REGION Network 5: 外呼下面有目标
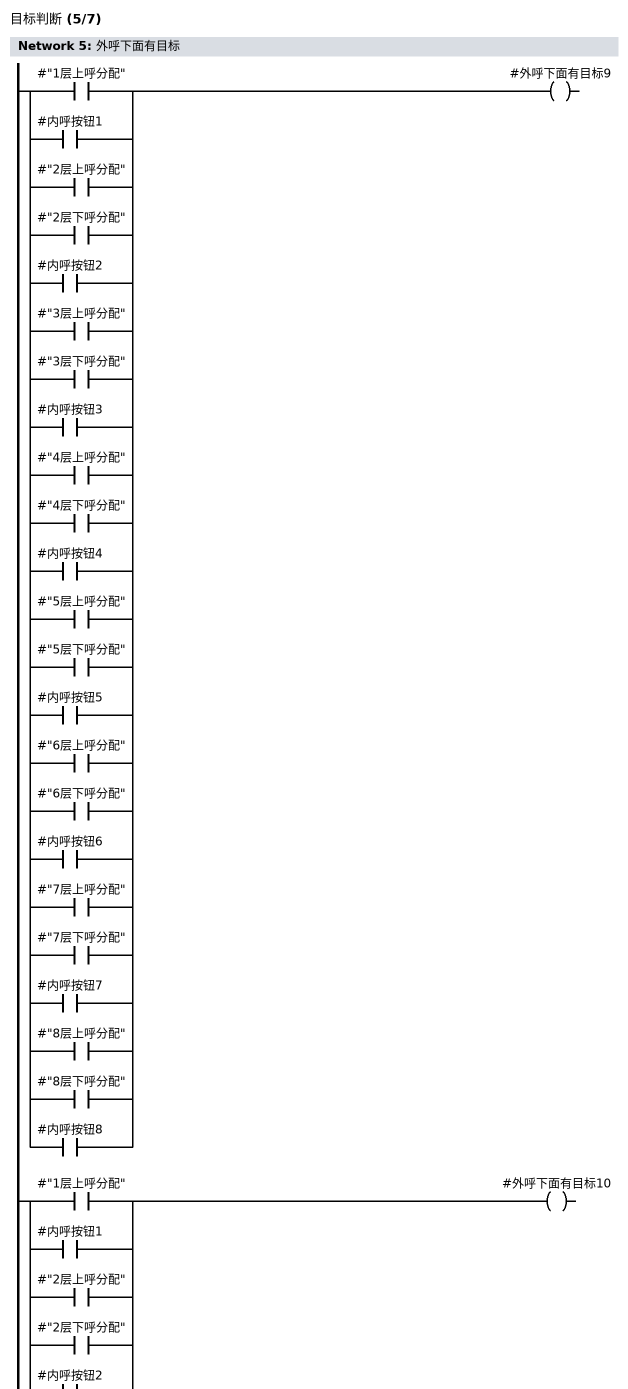
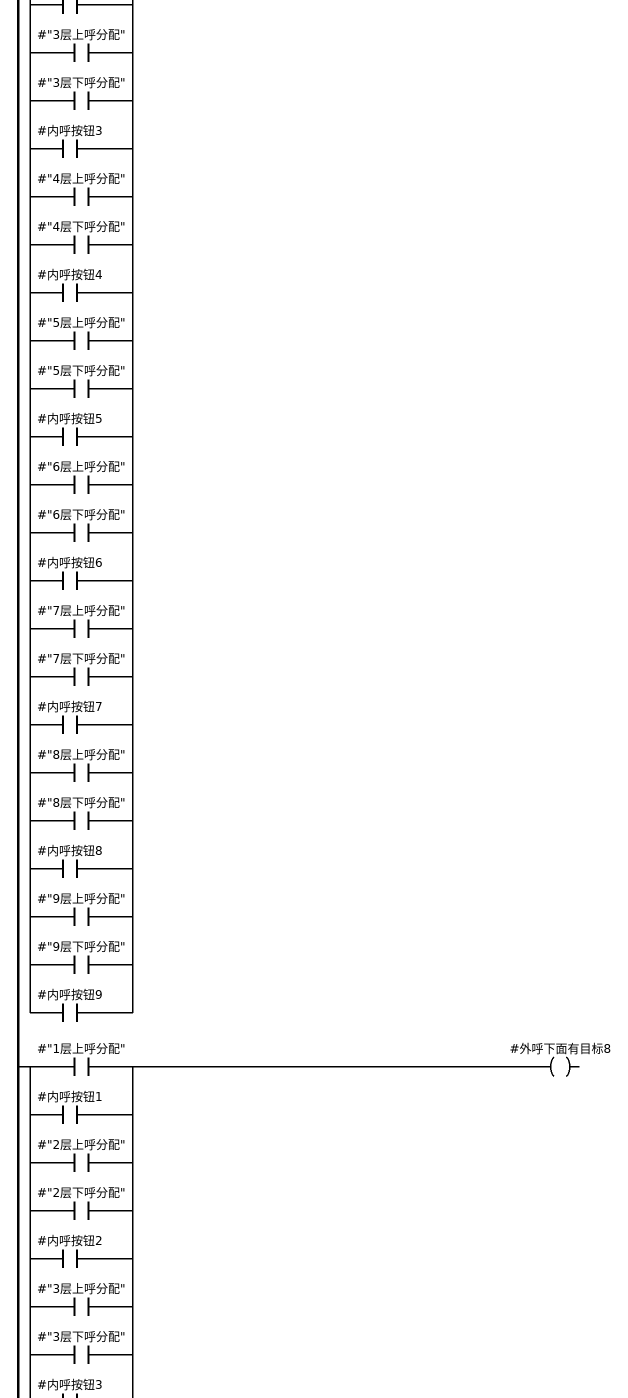
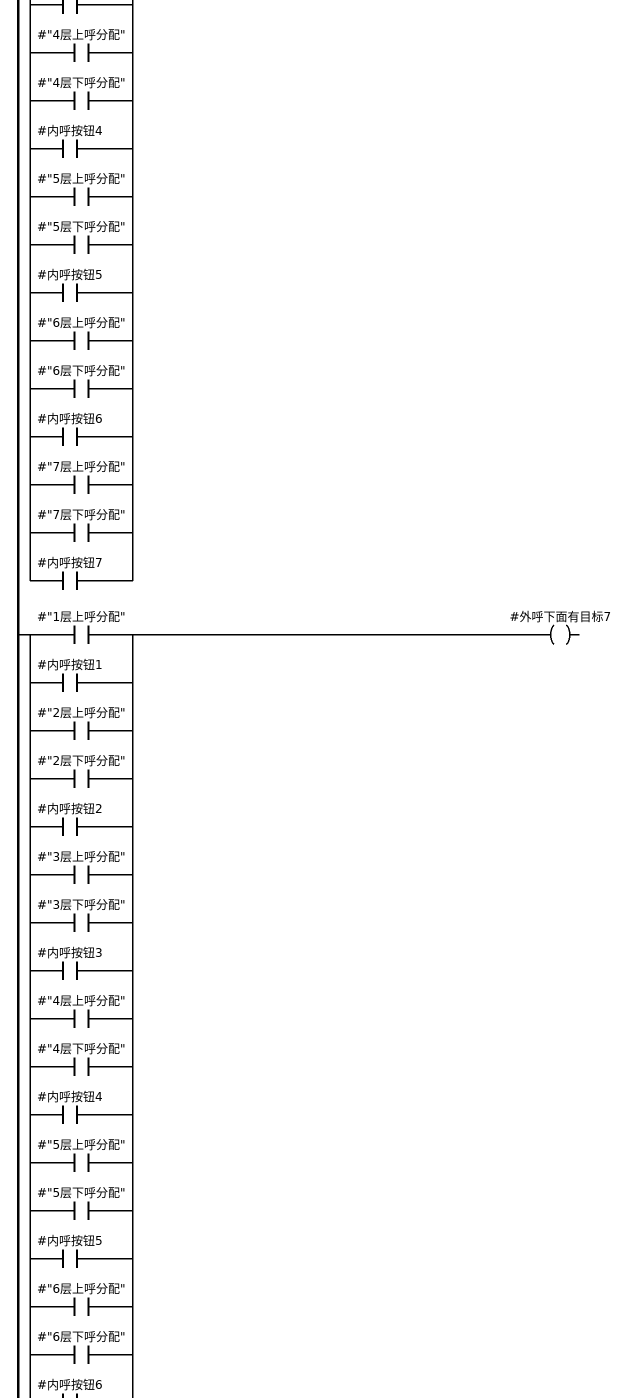
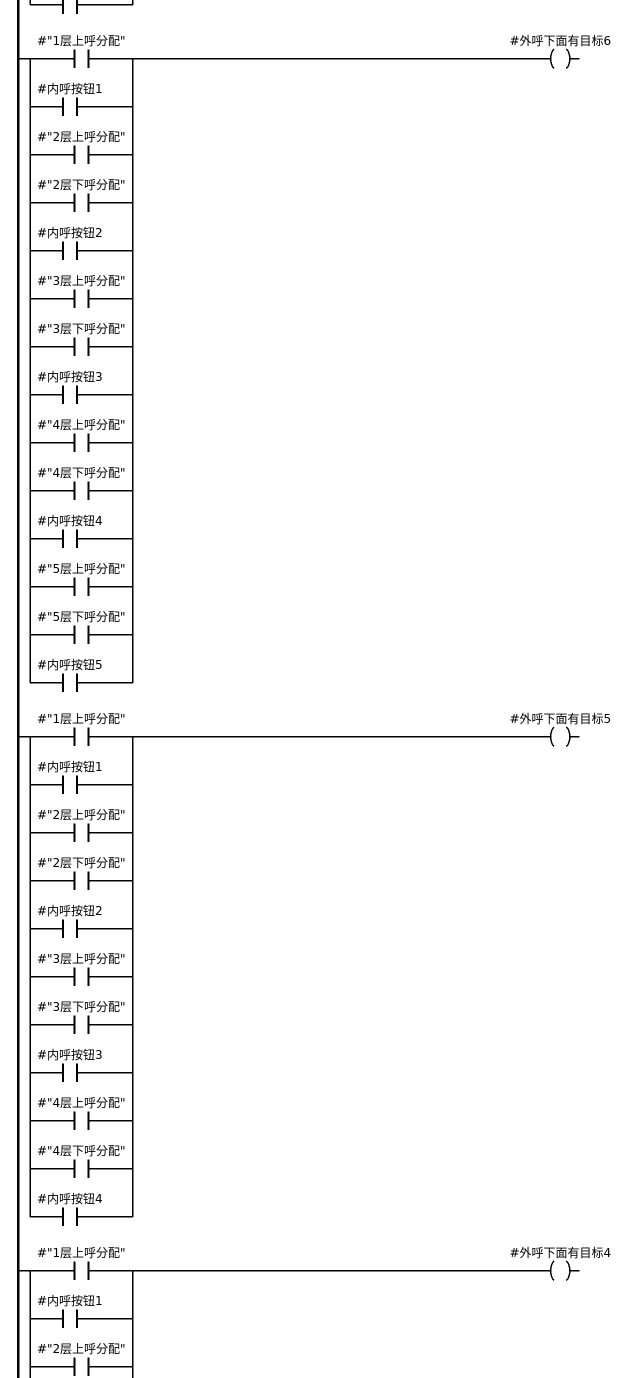
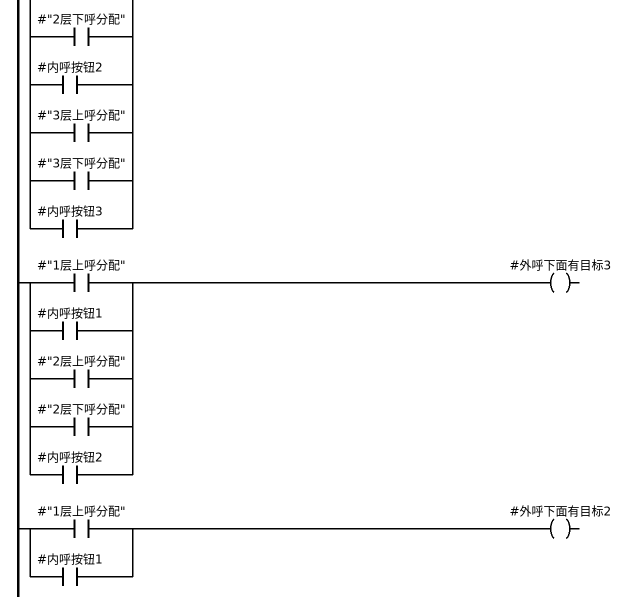
   RUNG wire#powerrail
      Contact( #"1层上呼分配" )
      wire#w1
      Coil( #外呼下面有目标9 )
   END_RUNG
   RUNG wire#powerrail
      Contact( #内呼按钮1 )
   END_RUNG wire#w1
   RUNG wire#powerrail
      Contact( #"2层上呼分配" )
   END_RUNG wire#w1
   RUNG wire#powerrail
      Contact( #"2层下呼分配" )
   END_RUNG wire#w1
   RUNG wire#powerrail
      Contact( #内呼按钮2 )
   END_RUNG wire#w1
   RUNG wire#powerrail
      Contact( #"3层上呼分配" )
   END_RUNG wire#w1
   RUNG wire#powerrail
      Contact( #"3层下呼分配" )
   END_RUNG wire#w1
   RUNG wire#powerrail
      Contact( #内呼按钮3 )
   END_RUNG wire#w1
   RUNG wire#powerrail
      Contact( #"4层上呼分配" )
   END_RUNG wire#w1
   RUNG wire#powerrail
      Contact( #"4层下呼分配" )
   END_RUNG wire#w1
   RUNG wire#powerrail
      Contact( #内呼按钮4 )
   END_RUNG wire#w1
   RUNG wire#powerrail
      Contact( #"5层上呼分配" )
   END_RUNG wire#w1
   RUNG wire#powerrail
      Contact( #"5层下呼分配" )
   END_RUNG wire#w1
   RUNG wire#powerrail
      Contact( #内呼按钮5 )
   END_RUNG wire#w1
   RUNG wire#powerrail
      Contact( #"6层上呼分配" )
   END_RUNG wire#w1
   RUNG wire#powerrail
      Contact( #"6层下呼分配" )
   END_RUNG wire#w1
   RUNG wire#powerrail
      Contact( #内呼按钮6 )
   END_RUNG wire#w1
   RUNG wire#powerrail
      Contact( #"7层上呼分配" )
   END_RUNG wire#w1
   RUNG wire#powerrail
      Contact( #"7层下呼分配" )
   END_RUNG wire#w1
   RUNG wire#powerrail
      Contact( #内呼按钮7 )
   END_RUNG wire#w1
   RUNG wire#powerrail
      Contact( #"8层上呼分配" )
   END_RUNG wire#w1
   RUNG wire#powerrail
      Contact( #"8层下呼分配" )
   END_RUNG wire#w1
   RUNG wire#powerrail
      Contact( #内呼按钮8 )
   END_RUNG wire#w1
   RUNG wire#powerrail
      Contact( #"1层上呼分配" )
      wire#w2
      Coil( #外呼下面有目标10 )
   END_RUNG
   RUNG wire#powerrail
      Contact( #内呼按钮1 )
   END_RUNG wire#w2
   RUNG wire#powerrail
      Contact( #"2层上呼分配" )
   END_RUNG wire#w2
   RUNG wire#powerrail
      Contact( #"2层下呼分配" )
   END_RUNG wire#w2
   RUNG wire#powerrail
      Contact( #内呼按钮2 )
   END_RUNG wire#w2
   RUNG wire#powerrail
      Contact( #"3层上呼分配" )
   END_RUNG wire#w2
   RUNG wire#powerrail
      Contact( #"3层下呼分配" )
   END_RUNG wire#w2
   RUNG wire#powerrail
      Contact( #内呼按钮3 )
   END_RUNG wire#w2
   RUNG wire#powerrail
      Contact( #"4层上呼分配" )
   END_RUNG wire#w2
   RUNG wire#powerrail
      Contact( #"4层下呼分配" )
   END_RUNG wire#w2
   RUNG wire#powerrail
      Contact( #内呼按钮4 )
   END_RUNG wire#w2
   RUNG wire#powerrail
      Contact( #"5层上呼分配" )
   END_RUNG wire#w2
   RUNG wire#powerrail
      Contact( #"5层下呼分配" )
   END_RUNG wire#w2
   RUNG wire#powerrail
      Contact( #内呼按钮5 )
   END_RUNG wire#w2
   RUNG wire#powerrail
      Contact( #"6层上呼分配" )
   END_RUNG wire#w2
   RUNG wire#powerrail
      Contact( #"6层下呼分配" )
   END_RUNG wire#w2
   RUNG wire#powerrail
      Contact( #内呼按钮6 )
   END_RUNG wire#w2
   RUNG wire#powerrail
      Contact( #"7层上呼分配" )
   END_RUNG wire#w2
   RUNG wire#powerrail
      Contact( #"7层下呼分配" )
   END_RUNG wire#w2
   RUNG wire#powerrail
      Contact( #内呼按钮7 )
   END_RUNG wire#w2
   RUNG wire#powerrail
      Contact( #"8层上呼分配" )
   END_RUNG wire#w2
   RUNG wire#powerrail
      Contact( #"8层下呼分配" )
   END_RUNG wire#w2
   RUNG wire#powerrail
      Contact( #内呼按钮8 )
   END_RUNG wire#w2
   RUNG wire#powerrail
      Contact( #"9层上呼分配" )
   END_RUNG wire#w2
   RUNG wire#powerrail
      Contact( #"9层下呼分配" )
   END_RUNG wire#w2
   RUNG wire#powerrail
      Contact( #内呼按钮9 )
   END_RUNG wire#w2
   RUNG wire#powerrail
      Contact( #"1层上呼分配" )
      wire#w3
      Coil( #外呼下面有目标8 )
   END_RUNG
   RUNG wire#powerrail
      Contact( #内呼按钮1 )
   END_RUNG wire#w3
   RUNG wire#powerrail
      Contact( #"2层上呼分配" )
   END_RUNG wire#w3
   RUNG wire#powerrail
      Contact( #"2层下呼分配" )
   END_RUNG wire#w3
   RUNG wire#powerrail
      Contact( #内呼按钮2 )
   END_RUNG wire#w3
   RUNG wire#powerrail
      Contact( #"3层上呼分配" )
   END_RUNG wire#w3
   RUNG wire#powerrail
      Contact( #"3层下呼分配" )
   END_RUNG wire#w3
   RUNG wire#powerrail
      Contact( #内呼按钮3 )
   END_RUNG wire#w3
   RUNG wire#powerrail
      Contact( #"4层上呼分配" )
   END_RUNG wire#w3
   RUNG wire#powerrail
      Contact( #"4层下呼分配" )
   END_RUNG wire#w3
   RUNG wire#powerrail
      Contact( #内呼按钮4 )
   END_RUNG wire#w3
   RUNG wire#powerrail
      Contact( #"5层上呼分配" )
   END_RUNG wire#w3
   RUNG wire#powerrail
      Contact( #"5层下呼分配" )
   END_RUNG wire#w3
   RUNG wire#powerrail
      Contact( #内呼按钮5 )
   END_RUNG wire#w3
   RUNG wire#powerrail
      Contact( #"6层上呼分配" )
   END_RUNG wire#w3
   RUNG wire#powerrail
      Contact( #"6层下呼分配" )
   END_RUNG wire#w3
   RUNG wire#powerrail
      Contact( #内呼按钮6 )
   END_RUNG wire#w3
   RUNG wire#powerrail
      Contact( #"7层上呼分配" )
   END_RUNG wire#w3
   RUNG wire#powerrail
      Contact( #"7层下呼分配" )
   END_RUNG wire#w3
   RUNG wire#powerrail
      Contact( #内呼按钮7 )
   END_RUNG wire#w3
   RUNG wire#powerrail
      Contact( #"1层上呼分配" )
      wire#w4
      Coil( #外呼下面有目标7 )
   END_RUNG
   RUNG wire#powerrail
      Contact( #内呼按钮1 )
   END_RUNG wire#w4
   RUNG wire#powerrail
      Contact( #"2层上呼分配" )
   END_RUNG wire#w4
   RUNG wire#powerrail
      Contact( #"2层下呼分配" )
   END_RUNG wire#w4
   RUNG wire#powerrail
      Contact( #内呼按钮2 )
   END_RUNG wire#w4
   RUNG wire#powerrail
      Contact( #"3层上呼分配" )
   END_RUNG wire#w4
   RUNG wire#powerrail
      Contact( #"3层下呼分配" )
   END_RUNG wire#w4
   RUNG wire#powerrail
      Contact( #内呼按钮3 )
   END_RUNG wire#w4
   RUNG wire#powerrail
      Contact( #"4层上呼分配" )
   END_RUNG wire#w4
   RUNG wire#powerrail
      Contact( #"4层下呼分配" )
   END_RUNG wire#w4
   RUNG wire#powerrail
      Contact( #内呼按钮4 )
   END_RUNG wire#w4
   RUNG wire#powerrail
      Contact( #"5层上呼分配" )
   END_RUNG wire#w4
   RUNG wire#powerrail
      Contact( #"5层下呼分配" )
   END_RUNG wire#w4
   RUNG wire#powerrail
      Contact( #内呼按钮5 )
   END_RUNG wire#w4
   RUNG wire#powerrail
      Contact( #"6层上呼分配" )
   END_RUNG wire#w4
   RUNG wire#powerrail
      Contact( #"6层下呼分配" )
   END_RUNG wire#w4
   RUNG wire#powerrail
      Contact( #内呼按钮6 )
   END_RUNG wire#w4
   RUNG wire#powerrail
      Contact( #"1层上呼分配" )
      wire#w5
      Coil( #外呼下面有目标6 )
   END_RUNG
   RUNG wire#powerrail
      Contact( #内呼按钮1 )
   END_RUNG wire#w5
   RUNG wire#powerrail
      Contact( #"2层上呼分配" )
   END_RUNG wire#w5
   RUNG wire#powerrail
      Contact( #"2层下呼分配" )
   END_RUNG wire#w5
   RUNG wire#powerrail
      Contact( #内呼按钮2 )
   END_RUNG wire#w5
   RUNG wire#powerrail
      Contact( #"3层上呼分配" )
   END_RUNG wire#w5
   RUNG wire#powerrail
      Contact( #"3层下呼分配" )
   END_RUNG wire#w5
   RUNG wire#powerrail
      Contact( #内呼按钮3 )
   END_RUNG wire#w5
   RUNG wire#powerrail
      Contact( #"4层上呼分配" )
   END_RUNG wire#w5
   RUNG wire#powerrail
      Contact( #"4层下呼分配" )
   END_RUNG wire#w5
   RUNG wire#powerrail
      Contact( #内呼按钮4 )
   END_RUNG wire#w5
   RUNG wire#powerrail
      Contact( #"5层上呼分配" )
   END_RUNG wire#w5
   RUNG wire#powerrail
      Contact( #"5层下呼分配" )
   END_RUNG wire#w5
   RUNG wire#powerrail
      Contact( #内呼按钮5 )
   END_RUNG wire#w5
   RUNG wire#powerrail
      Contact( #"1层上呼分配" )
      wire#w6
      Coil( #外呼下面有目标5 )
   END_RUNG
   RUNG wire#powerrail
      Contact( #内呼按钮1 )
   END_RUNG wire#w6
   RUNG wire#powerrail
      Contact( #"2层上呼分配" )
   END_RUNG wire#w6
   RUNG wire#powerrail
      Contact( #"2层下呼分配" )
   END_RUNG wire#w6
   RUNG wire#powerrail
      Contact( #内呼按钮2 )
   END_RUNG wire#w6
   RUNG wire#powerrail
      Contact( #"3层上呼分配" )
   END_RUNG wire#w6
   RUNG wire#powerrail
      Contact( #"3层下呼分配" )
   END_RUNG wire#w6
   RUNG wire#powerrail
      Contact( #内呼按钮3 )
   END_RUNG wire#w6
   RUNG wire#powerrail
      Contact( #"4层上呼分配" )
   END_RUNG wire#w6
   RUNG wire#powerrail
      Contact( #"4层下呼分配" )
   END_RUNG wire#w6
   RUNG wire#powerrail
      Contact( #内呼按钮4 )
   END_RUNG wire#w6
   RUNG wire#powerrail
      Contact( #"1层上呼分配" )
      wire#w7
      Coil( #外呼下面有目标4 )
   END_RUNG
   RUNG wire#powerrail
      Contact( #内呼按钮1 )
   END_RUNG wire#w7
   RUNG wire#powerrail
      Contact( #"2层上呼分配" )
   END_RUNG wire#w7
   RUNG wire#powerrail
      Contact( #"2层下呼分配" )
   END_RUNG wire#w7
   RUNG wire#powerrail
      Contact( #内呼按钮2 )
   END_RUNG wire#w7
   RUNG wire#powerrail
      Contact( #"3层上呼分配" )
   END_RUNG wire#w7
   RUNG wire#powerrail
      Contact( #"3层下呼分配" )
   END_RUNG wire#w7
   RUNG wire#powerrail
      Contact( #内呼按钮3 )
   END_RUNG wire#w7
   RUNG wire#powerrail
      Contact( #"1层上呼分配" )
      wire#w8
      Coil( #外呼下面有目标3 )
   END_RUNG
   RUNG wire#powerrail
      Contact( #内呼按钮1 )
   END_RUNG wire#w8
   RUNG wire#powerrail
      Contact( #"2层上呼分配" )
   END_RUNG wire#w8
   RUNG wire#powerrail
      Contact( #"2层下呼分配" )
   END_RUNG wire#w8
   RUNG wire#powerrail
      Contact( #内呼按钮2 )
   END_RUNG wire#w8
   RUNG wire#powerrail
      Contact( #"1层上呼分配" )
      wire#w9
      Coil( #外呼下面有目标2 )
   END_RUNG
   RUNG wire#powerrail
      Contact( #内呼按钮1 )
   END_RUNG wire#w9
   // the same network as SCL:
   #外呼下面有目标9 := #"1层上呼分配" OR #内呼按钮1 OR #"2层上呼分配" OR #"2层下呼分配" OR #内呼按钮2 OR #"3层上呼分配" OR #"3层下呼分配" OR #内呼按钮3 OR #"4层上呼分配" OR #"4层下呼分配" OR #内呼按钮4 OR #"5层上呼分配" OR #"5层下呼分配" OR #内呼按钮5 OR #"6层上呼分配" OR #"6层下呼分配" OR #内呼按钮6 OR #"7层上呼分配" OR #"7层下呼分配" OR #内呼按钮7 OR #"8层上呼分配" OR #"8层下呼分配" OR #内呼按钮8;
   #外呼下面有目标10 := #"1层上呼分配" OR #内呼按钮1 OR #"2层上呼分配" OR #"2层下呼分配" OR #内呼按钮2 OR #"3层上呼分配" OR #"3层下呼分配" OR #内呼按钮3 OR #"4层上呼分配" OR #"4层下呼分配" OR #内呼按钮4 OR #"5层上呼分配" OR #"5层下呼分配" OR #内呼按钮5 OR #"6层上呼分配" OR #"6层下呼分配" OR #内呼按钮6 OR #"7层上呼分配" OR #"7层下呼分配" OR #内呼按钮7 OR #"8层上呼分配" OR #"8层下呼分配" OR #内呼按钮8 OR #"9层上呼分配" OR #"9层下呼分配" OR #内呼按钮9;
   #外呼下面有目标8 := #"1层上呼分配" OR #内呼按钮1 OR #"2层上呼分配" OR #"2层下呼分配" OR #内呼按钮2 OR #"3层上呼分配" OR #"3层下呼分配" OR #内呼按钮3 OR #"4层上呼分配" OR #"4层下呼分配" OR #内呼按钮4 OR #"5层上呼分配" OR #"5层下呼分配" OR #内呼按钮5 OR #"6层上呼分配" OR #"6层下呼分配" OR #内呼按钮6 OR #"7层上呼分配" OR #"7层下呼分配" OR #内呼按钮7;
   #外呼下面有目标7 := #"1层上呼分配" OR #内呼按钮1 OR #"2层上呼分配" OR #"2层下呼分配" OR #内呼按钮2 OR #"3层上呼分配" OR #"3层下呼分配" OR #内呼按钮3 OR #"4层上呼分配" OR #"4层下呼分配" OR #内呼按钮4 OR #"5层上呼分配" OR #"5层下呼分配" OR #内呼按钮5 OR #"6层上呼分配" OR #"6层下呼分配" OR #内呼按钮6;
   #外呼下面有目标6 := #"1层上呼分配" OR #内呼按钮1 OR #"2层上呼分配" OR #"2层下呼分配" OR #内呼按钮2 OR #"3层上呼分配" OR #"3层下呼分配" OR #内呼按钮3 OR #"4层上呼分配" OR #"4层下呼分配" OR #内呼按钮4 OR #"5层上呼分配" OR #"5层下呼分配" OR #内呼按钮5;
   #外呼下面有目标5 := #"1层上呼分配" OR #内呼按钮1 OR #"2层上呼分配" OR #"2层下呼分配" OR #内呼按钮2 OR #"3层上呼分配" OR #"3层下呼分配" OR #内呼按钮3 OR #"4层上呼分配" OR #"4层下呼分配" OR #内呼按钮4;
   #外呼下面有目标4 := #"1层上呼分配" OR #内呼按钮1 OR #"2层上呼分配" OR #"2层下呼分配" OR #内呼按钮2 OR #"3层上呼分配" OR #"3层下呼分配" OR #内呼按钮3;
   #外呼下面有目标3 := #"1层上呼分配" OR #内呼按钮1 OR #"2层上呼分配" OR #"2层下呼分配" OR #内呼按钮2;
   #外呼下面有目标2 := #"1层上呼分配" OR #内呼按钮1;
END_REGION

REGION Network 6: 外呼上面有目标选取最远目标
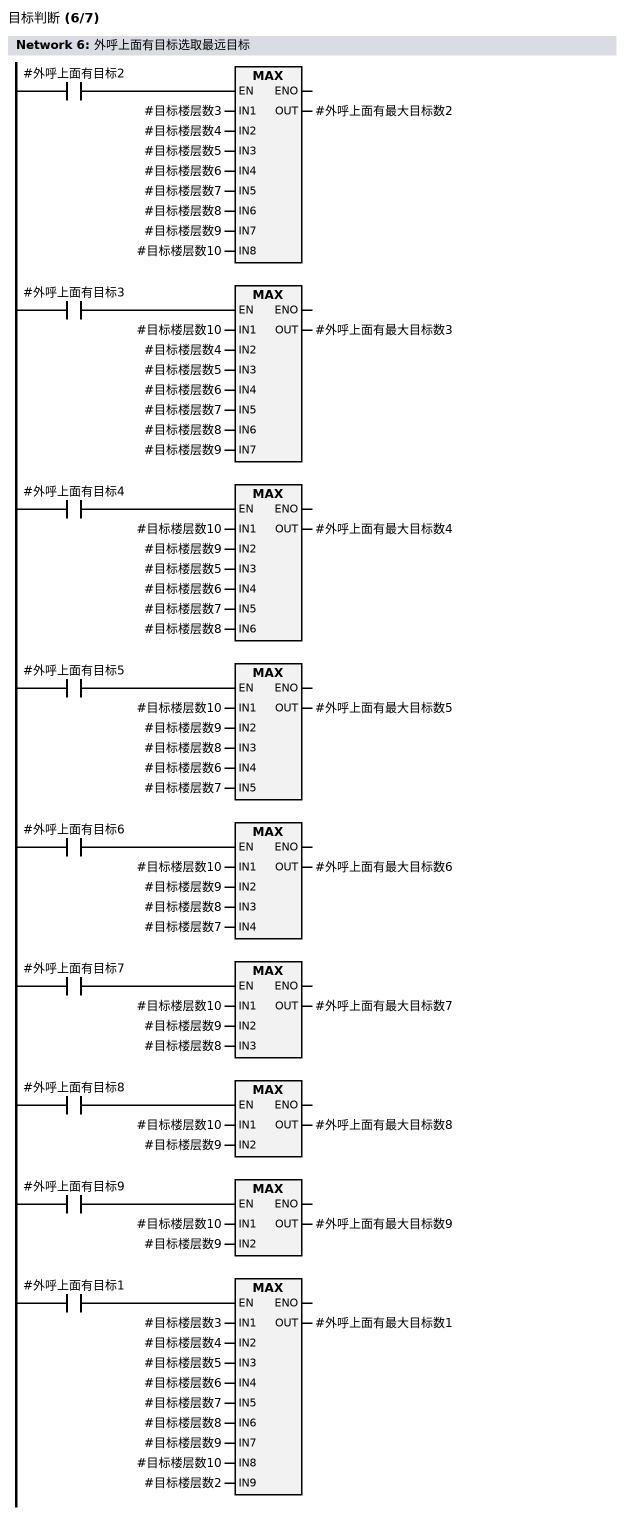
   IF #外呼上面有目标2 THEN
       #外呼上面有最大目标数2 := MAX(IN1 := #目标楼层数3, IN2 := #目标楼层数4, IN3 := #目标楼层数5, IN4 := #目标楼层数6, IN5 := #目标楼层数7, IN6 := #目标楼层数8, IN7 := #目标楼层数9, IN8 := #目标楼层数10);
   END_IF;
   IF #外呼上面有目标3 THEN
       #外呼上面有最大目标数3 := MAX(IN1 := #目标楼层数10, IN2 := #目标楼层数4, IN3 := #目标楼层数5, IN4 := #目标楼层数6, IN5 := #目标楼层数7, IN6 := #目标楼层数8, IN7 := #目标楼层数9);
   END_IF;
   IF #外呼上面有目标4 THEN
       #外呼上面有最大目标数4 := MAX(IN1 := #目标楼层数10, IN2 := #目标楼层数9, IN3 := #目标楼层数5, IN4 := #目标楼层数6, IN5 := #目标楼层数7, IN6 := #目标楼层数8);
   END_IF;
   IF #外呼上面有目标5 THEN
       #外呼上面有最大目标数5 := MAX(IN1 := #目标楼层数10, IN2 := #目标楼层数9, IN3 := #目标楼层数8, IN4 := #目标楼层数6, IN5 := #目标楼层数7);
   END_IF;
   IF #外呼上面有目标6 THEN
       #外呼上面有最大目标数6 := MAX(IN1 := #目标楼层数10, IN2 := #目标楼层数9, IN3 := #目标楼层数8, IN4 := #目标楼层数7);
   END_IF;
   IF #外呼上面有目标7 THEN #外呼上面有最大目标数7 := MAX(IN1 := #目标楼层数10, IN2 := #目标楼层数9, IN3 := #目标楼层数8); END_IF;
   IF #外呼上面有目标8 THEN #外呼上面有最大目标数8 := MAX(IN1 := #目标楼层数10, IN2 := #目标楼层数9); END_IF;
   IF #外呼上面有目标9 THEN #外呼上面有最大目标数9 := MAX(IN1 := #目标楼层数10, IN2 := #目标楼层数9); END_IF;
   IF #外呼上面有目标1 THEN
       #外呼上面有最大目标数1 := MAX(IN1 := #目标楼层数3, IN2 := #目标楼层数4, IN3 := #目标楼层数5, IN4 := #目标楼层数6, IN5 := #目标楼层数7, IN6 := #目标楼层数8, IN7 := #目标楼层数9, IN8 := #目标楼层数10, IN9 := #目标楼层数2);
   END_IF;
END_REGION

REGION Network 7: 外呼下面有目标选取最远目标
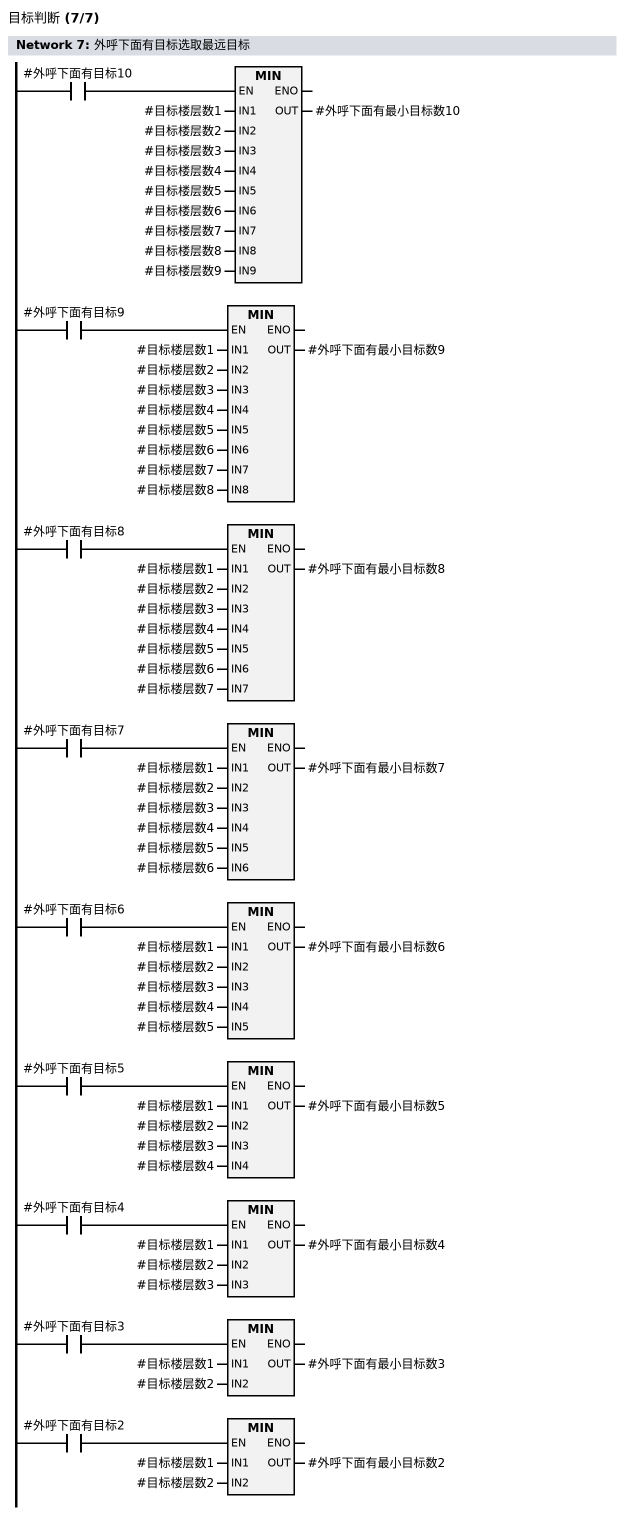
   IF #外呼下面有目标10 THEN
       #外呼下面有最小目标数10 := MIN(IN1 := #目标楼层数1, IN2 := #目标楼层数2, IN3 := #目标楼层数3, IN4 := #目标楼层数4, IN5 := #目标楼层数5, IN6 := #目标楼层数6, IN7 := #目标楼层数7, IN8 := #目标楼层数8, IN9 := #目标楼层数9);
   END_IF;
   IF #外呼下面有目标9 THEN
       #外呼下面有最小目标数9 := MIN(IN1 := #目标楼层数1, IN2 := #目标楼层数2, IN3 := #目标楼层数3, IN4 := #目标楼层数4, IN5 := #目标楼层数5, IN6 := #目标楼层数6, IN7 := #目标楼层数7, IN8 := #目标楼层数8);
   END_IF;
   IF #外呼下面有目标8 THEN
       #外呼下面有最小目标数8 := MIN(IN1 := #目标楼层数1, IN2 := #目标楼层数2, IN3 := #目标楼层数3, IN4 := #目标楼层数4, IN5 := #目标楼层数5, IN6 := #目标楼层数6, IN7 := #目标楼层数7);
   END_IF;
   IF #外呼下面有目标7 THEN
       #外呼下面有最小目标数7 := MIN(IN1 := #目标楼层数1, IN2 := #目标楼层数2, IN3 := #目标楼层数3, IN4 := #目标楼层数4, IN5 := #目标楼层数5, IN6 := #目标楼层数6);
   END_IF;
   IF #外呼下面有目标6 THEN
       #外呼下面有最小目标数6 := MIN(IN1 := #目标楼层数1, IN2 := #目标楼层数2, IN3 := #目标楼层数3, IN4 := #目标楼层数4, IN5 := #目标楼层数5);
   END_IF;
   IF #外呼下面有目标5 THEN
       #外呼下面有最小目标数5 := MIN(IN1 := #目标楼层数1, IN2 := #目标楼层数2, IN3 := #目标楼层数3, IN4 := #目标楼层数4);
   END_IF;
   IF #外呼下面有目标4 THEN #外呼下面有最小目标数4 := MIN(IN1 := #目标楼层数1, IN2 := #目标楼层数2, IN3 := #目标楼层数3); END_IF;
   IF #外呼下面有目标3 THEN #外呼下面有最小目标数3 := MIN(IN1 := #目标楼层数1, IN2 := #目标楼层数2); END_IF;
   IF #外呼下面有目标2 THEN #外呼下面有最小目标数2 := MIN(IN1 := #目标楼层数1, IN2 := #目标楼层数2); END_IF;
END_REGION
END_FUNCTION_BLOCK

FUNCTION_BLOCK "初始化低速模式"   // FB4, LAD
{ S7_Optimized_Access := 'TRUE' }
VERSION : 0.1
   VAR_INPUT
      当前楼层数 : Int;
      初始化低速运行 : Bool;
      "1层上行呼梯按钮指示灯" : Bool;
      "2层上行呼梯按钮指示灯" : Bool;
      "3层上行呼梯按钮指示灯" : Bool;
      "4层上行呼梯按钮指示灯" : Bool;
      "5层上行呼梯按钮指示灯" : Bool;
      "6层上行呼梯按钮指示灯" : Bool;
      "7层上行呼梯按钮指示灯" : Bool;
      "8层上行呼梯按钮指示灯" : Bool;
      "9层上行呼梯按钮指示灯" : Bool;
      "2层下行呼梯按钮指示灯" : Bool;
      "3层下行呼梯按钮指示灯" : Bool;
      "4层下行呼梯按钮指示灯" : Bool;
      "5层下行呼梯按钮指示灯" : Bool;
      "6层下行呼梯按钮指示灯" : Bool;
      "7层下行呼梯按钮指示灯" : Bool;
      "8层下行呼梯按钮指示灯" : Bool;
      "9层下行呼梯按钮指示灯" : Bool;
      "10层下行呼梯按钮指示灯" : Bool;
      "1号梯1层按钮指示灯" : Bool;
      "1号梯2层按钮指示灯" : Bool;
      "1号梯3层按钮指示灯" : Bool;
      "1号梯4层按钮指示灯" : Bool;
      "1号梯5层按钮指示灯" : Bool;
      "1号梯6层按钮指示灯" : Bool;
      "1号梯7层按钮指示灯" : Bool;
      "1号梯8层按钮指示灯" : Bool;
      "1号梯9层按钮指示灯" : Bool;
      "1号梯10层按钮指示灯" : Bool;
      正处于故障中 : Bool;
      "存在安全隐患（光幕）" : Bool;
      置0为完成开门 : Bool;
      置0为完成关门 : Bool;
      "1号梯上行指示" : Bool;
      "1号梯下行指示" : Bool;
      "1号梯检修信号" : Bool;
      "1号梯上行接触器" : Bool;
      "1号梯下行接触器" : Bool;
      "1号梯外呼上面无目标2" : Bool;
      "1号梯外呼上面无目标3" : Bool;
      "1号梯外呼上面无目标4" : Bool;
      "1号梯外呼上面无目标5" : Bool;
      "1号梯外呼上面无目标6" : Bool;
      "1号梯外呼上面无目标7" : Bool;
      "1号梯外呼上面无目标8" : Bool;
      "1号梯外呼上面无目标9" : Bool;
      "1号梯外呼下面无目标2" : Bool;
      "1号梯外呼下面无目标3" : Bool;
      "1号梯外呼下面无目标4" : Bool;
      "1号梯外呼下面无目标5" : Bool;
      "1号梯外呼下面无目标6" : Bool;
      "1号梯外呼下面无目标7" : Bool;
      "1号梯外呼下面无目标8" : Bool;
      "1号梯外呼下面无目标9" : Bool;
   END_VAR
   VAR_OUTPUT
      "1号梯高速接触器" : Bool;
      将要停梯 : Bool;
      "1号梯低速接触器" : Bool;
   END_VAR
   VAR
      "1楼相关" : Bool;
      "2楼相关" : Bool;
      "3楼相关" : Bool;
      "4楼相关" : Bool;
      "5楼相关" : Bool;
      "6楼相关" : Bool;
      "7楼相关" : Bool;
      "8楼相关" : Bool;
      "9楼相关" : Bool;
      "10楼相关" : Bool;
      分类上行特殊 : Bool;
      分类下行特殊 : Bool;
      中间变量1 : Bool;
      中间变量2 : Bool;
      中间变量3 : Bool;
      中间变量4 : Bool;
      中间变量5 : Bool;
      中间变量6 : Bool;
      中间变量7 : Bool;
   END_VAR
BEGIN

REGION Network 1: 低速上下行（前正常指令，后最后指令）
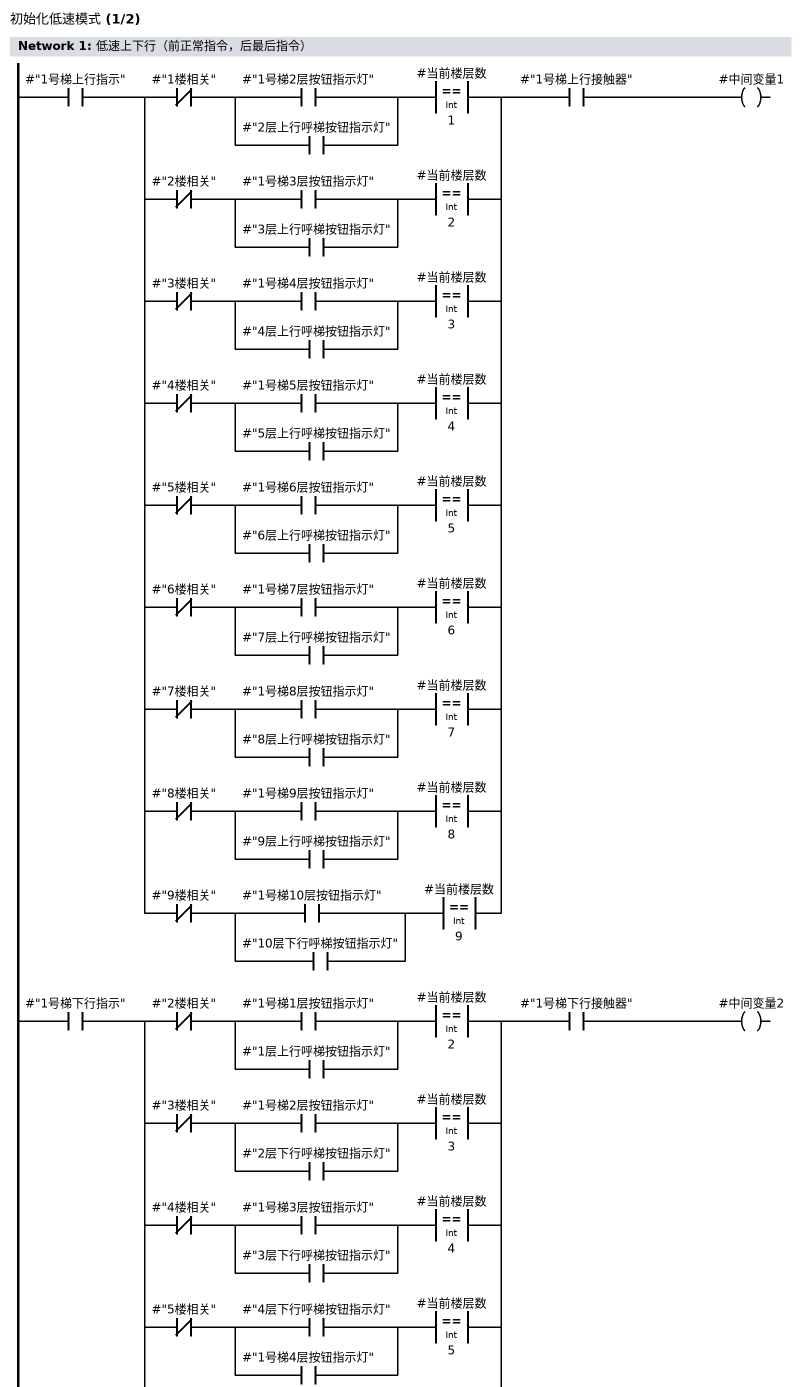
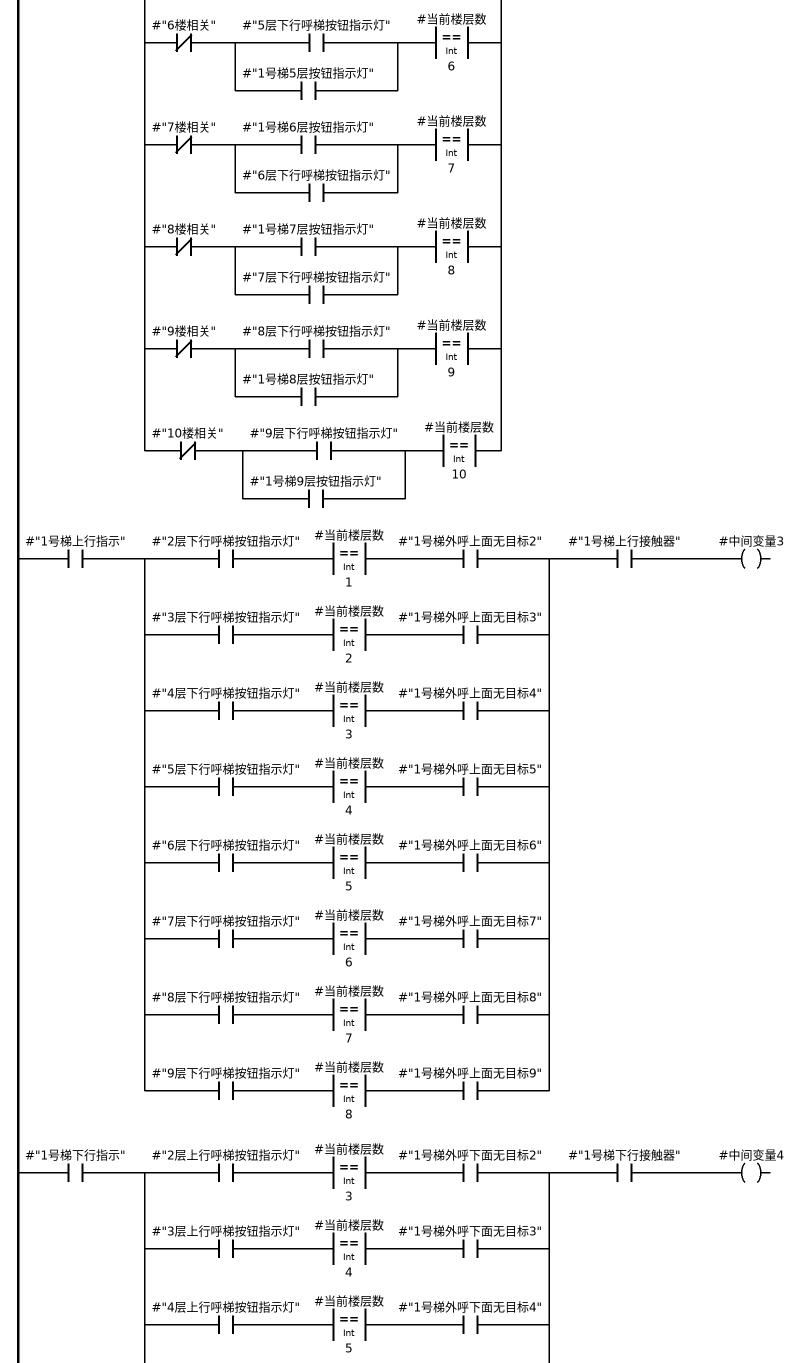
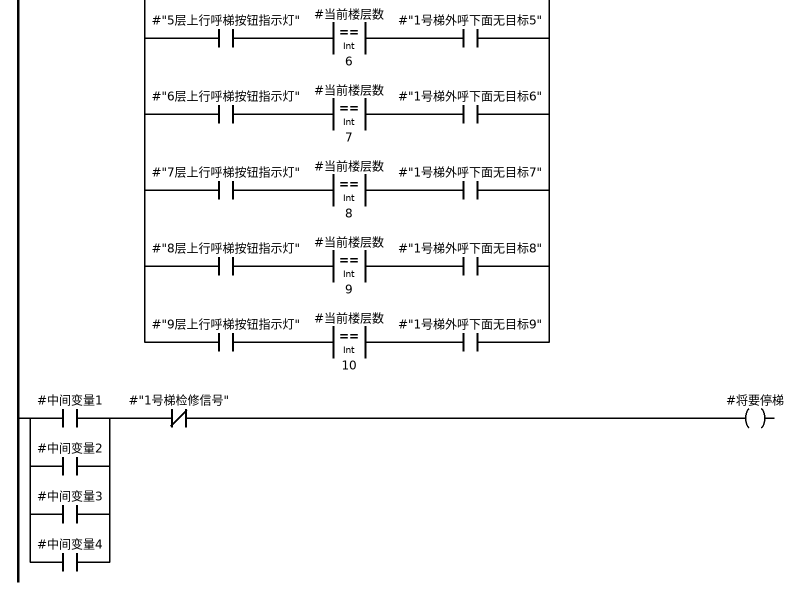
   RUNG wire#powerrail
      Contact( #"1号梯上行指示" )
      wire#w1
      I_Contact( #"1楼相关" )
      wire#w2
      Contact( #"1号梯2层按钮指示灯" )
      wire#w3
      { S7_Templates := "SrcType := Int" } EQ_Contact(in1 := #当前楼层数, in2 := 1)
      wire#w4
      Contact( #"1号梯上行接触器" )
      Coil( #中间变量1 )
   END_RUNG
   RUNG wire#w2
      Contact( #"2层上行呼梯按钮指示灯" )
   END_RUNG wire#w3
   RUNG wire#w1
      I_Contact( #"2楼相关" )
      wire#w5
      Contact( #"1号梯3层按钮指示灯" )
      wire#w6
      { S7_Templates := "SrcType := Int" } EQ_Contact(in1 := #当前楼层数, in2 := 2)
   END_RUNG wire#w4
   RUNG wire#w5
      Contact( #"3层上行呼梯按钮指示灯" )
   END_RUNG wire#w6
   RUNG wire#w1
      I_Contact( #"3楼相关" )
      wire#w7
      Contact( #"1号梯4层按钮指示灯" )
      wire#w8
      { S7_Templates := "SrcType := Int" } EQ_Contact(in1 := #当前楼层数, in2 := 3)
   END_RUNG wire#w4
   RUNG wire#w7
      Contact( #"4层上行呼梯按钮指示灯" )
   END_RUNG wire#w8
   RUNG wire#w1
      I_Contact( #"4楼相关" )
      wire#w9
      Contact( #"1号梯5层按钮指示灯" )
      wire#w10
      { S7_Templates := "SrcType := Int" } EQ_Contact(in1 := #当前楼层数, in2 := 4)
   END_RUNG wire#w4
   RUNG wire#w9
      Contact( #"5层上行呼梯按钮指示灯" )
   END_RUNG wire#w10
   RUNG wire#w1
      I_Contact( #"5楼相关" )
      wire#w11
      Contact( #"1号梯6层按钮指示灯" )
      wire#w12
      { S7_Templates := "SrcType := Int" } EQ_Contact(in1 := #当前楼层数, in2 := 5)
   END_RUNG wire#w4
   RUNG wire#w11
      Contact( #"6层上行呼梯按钮指示灯" )
   END_RUNG wire#w12
   RUNG wire#w1
      I_Contact( #"6楼相关" )
      wire#w13
      Contact( #"1号梯7层按钮指示灯" )
      wire#w14
      { S7_Templates := "SrcType := Int" } EQ_Contact(in1 := #当前楼层数, in2 := 6)
   END_RUNG wire#w4
   RUNG wire#w13
      Contact( #"7层上行呼梯按钮指示灯" )
   END_RUNG wire#w14
   RUNG wire#w1
      I_Contact( #"7楼相关" )
      wire#w15
      Contact( #"1号梯8层按钮指示灯" )
      wire#w16
      { S7_Templates := "SrcType := Int" } EQ_Contact(in1 := #当前楼层数, in2 := 7)
   END_RUNG wire#w4
   RUNG wire#w15
      Contact( #"8层上行呼梯按钮指示灯" )
   END_RUNG wire#w16
   RUNG wire#w1
      I_Contact( #"8楼相关" )
      wire#w17
      Contact( #"1号梯9层按钮指示灯" )
      wire#w18
      { S7_Templates := "SrcType := Int" } EQ_Contact(in1 := #当前楼层数, in2 := 8)
   END_RUNG wire#w4
   RUNG wire#w17
      Contact( #"9层上行呼梯按钮指示灯" )
   END_RUNG wire#w18
   RUNG wire#w1
      I_Contact( #"9楼相关" )
      wire#w19
      Contact( #"1号梯10层按钮指示灯" )
      wire#w20
      { S7_Templates := "SrcType := Int" } EQ_Contact(in1 := #当前楼层数, in2 := 9)
   END_RUNG wire#w4
   RUNG wire#w19
      Contact( #"10层下行呼梯按钮指示灯" )
   END_RUNG wire#w20
   RUNG wire#powerrail
      Contact( #"1号梯下行指示" )
      wire#w21
      I_Contact( #"2楼相关" )
      wire#w22
      Contact( #"1号梯1层按钮指示灯" )
      wire#w23
      { S7_Templates := "SrcType := Int" } EQ_Contact(in1 := #当前楼层数, in2 := 2)
      wire#w24
      Contact( #"1号梯下行接触器" )
      Coil( #中间变量2 )
   END_RUNG
   RUNG wire#w22
      Contact( #"1层上行呼梯按钮指示灯" )
   END_RUNG wire#w23
   RUNG wire#w21
      I_Contact( #"3楼相关" )
      wire#w25
      Contact( #"1号梯2层按钮指示灯" )
      wire#w26
      { S7_Templates := "SrcType := Int" } EQ_Contact(in1 := #当前楼层数, in2 := 3)
   END_RUNG wire#w24
   RUNG wire#w25
      Contact( #"2层下行呼梯按钮指示灯" )
   END_RUNG wire#w26
   RUNG wire#w21
      I_Contact( #"4楼相关" )
      wire#w27
      Contact( #"1号梯3层按钮指示灯" )
      wire#w28
      { S7_Templates := "SrcType := Int" } EQ_Contact(in1 := #当前楼层数, in2 := 4)
   END_RUNG wire#w24
   RUNG wire#w27
      Contact( #"3层下行呼梯按钮指示灯" )
   END_RUNG wire#w28
   RUNG wire#w21
      I_Contact( #"5楼相关" )
      wire#w29
      Contact( #"4层下行呼梯按钮指示灯" )
      wire#w30
      { S7_Templates := "SrcType := Int" } EQ_Contact(in1 := #当前楼层数, in2 := 5)
   END_RUNG wire#w24
   RUNG wire#w29
      Contact( #"1号梯4层按钮指示灯" )
   END_RUNG wire#w30
   RUNG wire#w21
      I_Contact( #"6楼相关" )
      wire#w31
      Contact( #"5层下行呼梯按钮指示灯" )
      wire#w32
      { S7_Templates := "SrcType := Int" } EQ_Contact(in1 := #当前楼层数, in2 := 6)
   END_RUNG wire#w24
   RUNG wire#w31
      Contact( #"1号梯5层按钮指示灯" )
   END_RUNG wire#w32
   RUNG wire#w21
      I_Contact( #"7楼相关" )
      wire#w33
      Contact( #"1号梯6层按钮指示灯" )
      wire#w34
      { S7_Templates := "SrcType := Int" } EQ_Contact(in1 := #当前楼层数, in2 := 7)
   END_RUNG wire#w24
   RUNG wire#w33
      Contact( #"6层下行呼梯按钮指示灯" )
   END_RUNG wire#w34
   RUNG wire#w21
      I_Contact( #"8楼相关" )
      wire#w35
      Contact( #"1号梯7层按钮指示灯" )
      wire#w36
      { S7_Templates := "SrcType := Int" } EQ_Contact(in1 := #当前楼层数, in2 := 8)
   END_RUNG wire#w24
   RUNG wire#w35
      Contact( #"7层下行呼梯按钮指示灯" )
   END_RUNG wire#w36
   RUNG wire#w21
      I_Contact( #"9楼相关" )
      wire#w37
      Contact( #"8层下行呼梯按钮指示灯" )
      wire#w38
      { S7_Templates := "SrcType := Int" } EQ_Contact(in1 := #当前楼层数, in2 := 9)
   END_RUNG wire#w24
   RUNG wire#w37
      Contact( #"1号梯8层按钮指示灯" )
   END_RUNG wire#w38
   RUNG wire#w21
      I_Contact( #"10楼相关" )
      wire#w39
      Contact( #"9层下行呼梯按钮指示灯" )
      wire#w40
      { S7_Templates := "SrcType := Int" } EQ_Contact(in1 := #当前楼层数, in2 := 10)
   END_RUNG wire#w24
   RUNG wire#w39
      Contact( #"1号梯9层按钮指示灯" )
   END_RUNG wire#w40
   RUNG wire#powerrail
      Contact( #"1号梯上行指示" )
      wire#w41
      Contact( #"2层下行呼梯按钮指示灯" )
      { S7_Templates := "SrcType := Int" } EQ_Contact(in1 := #当前楼层数, in2 := 1)
      Contact( #"1号梯外呼上面无目标2" )
      wire#w42
      Contact( #"1号梯上行接触器" )
      Coil( #中间变量3 )
   END_RUNG
   RUNG wire#w41
      Contact( #"3层下行呼梯按钮指示灯" )
      { S7_Templates := "SrcType := Int" } EQ_Contact(in1 := #当前楼层数, in2 := 2)
      Contact( #"1号梯外呼上面无目标3" )
   END_RUNG wire#w42
   RUNG wire#w41
      Contact( #"4层下行呼梯按钮指示灯" )
      { S7_Templates := "SrcType := Int" } EQ_Contact(in1 := #当前楼层数, in2 := 3)
      Contact( #"1号梯外呼上面无目标4" )
   END_RUNG wire#w42
   RUNG wire#w41
      Contact( #"5层下行呼梯按钮指示灯" )
      { S7_Templates := "SrcType := Int" } EQ_Contact(in1 := #当前楼层数, in2 := 4)
      Contact( #"1号梯外呼上面无目标5" )
   END_RUNG wire#w42
   RUNG wire#w41
      Contact( #"6层下行呼梯按钮指示灯" )
      { S7_Templates := "SrcType := Int" } EQ_Contact(in1 := #当前楼层数, in2 := 5)
      Contact( #"1号梯外呼上面无目标6" )
   END_RUNG wire#w42
   RUNG wire#w41
      Contact( #"7层下行呼梯按钮指示灯" )
      { S7_Templates := "SrcType := Int" } EQ_Contact(in1 := #当前楼层数, in2 := 6)
      Contact( #"1号梯外呼上面无目标7" )
   END_RUNG wire#w42
   RUNG wire#w41
      Contact( #"8层下行呼梯按钮指示灯" )
      { S7_Templates := "SrcType := Int" } EQ_Contact(in1 := #当前楼层数, in2 := 7)
      Contact( #"1号梯外呼上面无目标8" )
   END_RUNG wire#w42
   RUNG wire#w41
      Contact( #"9层下行呼梯按钮指示灯" )
      { S7_Templates := "SrcType := Int" } EQ_Contact(in1 := #当前楼层数, in2 := 8)
      Contact( #"1号梯外呼上面无目标9" )
   END_RUNG wire#w42
   RUNG wire#powerrail
      Contact( #"1号梯下行指示" )
      wire#w43
      Contact( #"2层上行呼梯按钮指示灯" )
      { S7_Templates := "SrcType := Int" } EQ_Contact(in1 := #当前楼层数, in2 := 3)
      Contact( #"1号梯外呼下面无目标2" )
      wire#w44
      Contact( #"1号梯下行接触器" )
      Coil( #中间变量4 )
   END_RUNG
   RUNG wire#w43
      Contact( #"3层上行呼梯按钮指示灯" )
      { S7_Templates := "SrcType := Int" } EQ_Contact(in1 := #当前楼层数, in2 := 4)
      Contact( #"1号梯外呼下面无目标3" )
   END_RUNG wire#w44
   RUNG wire#w43
      Contact( #"4层上行呼梯按钮指示灯" )
      { S7_Templates := "SrcType := Int" } EQ_Contact(in1 := #当前楼层数, in2 := 5)
      Contact( #"1号梯外呼下面无目标4" )
   END_RUNG wire#w44
   RUNG wire#w43
      Contact( #"5层上行呼梯按钮指示灯" )
      { S7_Templates := "SrcType := Int" } EQ_Contact(in1 := #当前楼层数, in2 := 6)
      Contact( #"1号梯外呼下面无目标5" )
   END_RUNG wire#w44
   RUNG wire#w43
      Contact( #"6层上行呼梯按钮指示灯" )
      { S7_Templates := "SrcType := Int" } EQ_Contact(in1 := #当前楼层数, in2 := 7)
      Contact( #"1号梯外呼下面无目标6" )
   END_RUNG wire#w44
   RUNG wire#w43
      Contact( #"7层上行呼梯按钮指示灯" )
      { S7_Templates := "SrcType := Int" } EQ_Contact(in1 := #当前楼层数, in2 := 8)
      Contact( #"1号梯外呼下面无目标7" )
   END_RUNG wire#w44
   RUNG wire#w43
      Contact( #"8层上行呼梯按钮指示灯" )
      { S7_Templates := "SrcType := Int" } EQ_Contact(in1 := #当前楼层数, in2 := 9)
      Contact( #"1号梯外呼下面无目标8" )
   END_RUNG wire#w44
   RUNG wire#w43
      Contact( #"9层上行呼梯按钮指示灯" )
      { S7_Templates := "SrcType := Int" } EQ_Contact(in1 := #当前楼层数, in2 := 10)
      Contact( #"1号梯外呼下面无目标9" )
   END_RUNG wire#w44
   RUNG wire#powerrail
      Contact( #中间变量1 )
      wire#w45
      I_Contact( #"1号梯检修信号" )
      Coil( #将要停梯 )
   END_RUNG
   RUNG wire#powerrail
      Contact( #中间变量2 )
   END_RUNG wire#w45
   RUNG wire#powerrail
      Contact( #中间变量3 )
   END_RUNG wire#w45
   RUNG wire#powerrail
      Contact( #中间变量4 )
   END_RUNG wire#w45
   // the same network as SCL:
   #中间变量1 := #"1号梯上行指示" AND ((NOT #"1楼相关" AND (#"1号梯2层按钮指示灯" OR #"2层上行呼梯按钮指示灯") AND (#当前楼层数 = 1)) OR (NOT #"2楼相关" AND (#"1号梯3层按钮指示灯" OR #"3层上行呼梯按钮指示灯") AND (#当前楼层数 = 2)) OR (NOT #"3楼相关" AND (#"1号梯4层按钮指示灯" OR #"4层上行呼梯按钮指示灯") AND (#当前楼层数 = 3)) OR (NOT #"4楼相关" AND (#"1号梯5层按钮指示灯" OR #"5层上行呼梯按钮指示灯") AND (#当前楼层数 = 4)) OR (NOT #"5楼相关" AND (#"1号梯6层按钮指示灯" OR #"6层上行呼梯按钮指示灯") AND (#当前楼层数 = 5)) OR (NOT #"6楼相关" AND (#"1号梯7层按钮指示灯" OR #"7层上行呼梯按钮指示灯") AND (#当前楼层数 = 6)) OR (NOT #"7楼相关" AND (#"1号梯8层按钮指示灯" OR #"8层上行呼梯按钮指示灯") AND (#当前楼层数 = 7)) OR (NOT #"8楼相关" AND (#"1号梯9层按钮指示灯" OR #"9层上行呼梯按钮指示灯") AND (#当前楼层数 = 8)) OR (NOT #"9楼相关" AND (#"1号梯10层按钮指示灯" OR #"10层下行呼梯按钮指示灯") AND (#当前楼层数 = 9))) AND #"1号梯上行接触器";
   #中间变量2 := #"1号梯下行指示" AND ((NOT #"2楼相关" AND (#"1号梯1层按钮指示灯" OR #"1层上行呼梯按钮指示灯") AND (#当前楼层数 = 2)) OR (NOT #"3楼相关" AND (#"1号梯2层按钮指示灯" OR #"2层下行呼梯按钮指示灯") AND (#当前楼层数 = 3)) OR (NOT #"4楼相关" AND (#"1号梯3层按钮指示灯" OR #"3层下行呼梯按钮指示灯") AND (#当前楼层数 = 4)) OR (NOT #"5楼相关" AND (#"4层下行呼梯按钮指示灯" OR #"1号梯4层按钮指示灯") AND (#当前楼层数 = 5)) OR (NOT #"6楼相关" AND (#"5层下行呼梯按钮指示灯" OR #"1号梯5层按钮指示灯") AND (#当前楼层数 = 6)) OR (NOT #"7楼相关" AND (#"1号梯6层按钮指示灯" OR #"6层下行呼梯按钮指示灯") AND (#当前楼层数 = 7)) OR (NOT #"8楼相关" AND (#"1号梯7层按钮指示灯" OR #"7层下行呼梯按钮指示灯") AND (#当前楼层数 = 8)) OR (NOT #"9楼相关" AND (#"8层下行呼梯按钮指示灯" OR #"1号梯8层按钮指示灯") AND (#当前楼层数 = 9)) OR (NOT #"10楼相关" AND (#"9层下行呼梯按钮指示灯" OR #"1号梯9层按钮指示灯") AND (#当前楼层数 = 10))) AND #"1号梯下行接触器";
   #中间变量3 := #"1号梯上行指示" AND ((#"2层下行呼梯按钮指示灯" AND (#当前楼层数 = 1) AND #"1号梯外呼上面无目标2") OR (#"3层下行呼梯按钮指示灯" AND (#当前楼层数 = 2) AND #"1号梯外呼上面无目标3") OR (#"4层下行呼梯按钮指示灯" AND (#当前楼层数 = 3) AND #"1号梯外呼上面无目标4") OR (#"5层下行呼梯按钮指示灯" AND (#当前楼层数 = 4) AND #"1号梯外呼上面无目标5") OR (#"6层下行呼梯按钮指示灯" AND (#当前楼层数 = 5) AND #"1号梯外呼上面无目标6") OR (#"7层下行呼梯按钮指示灯" AND (#当前楼层数 = 6) AND #"1号梯外呼上面无目标7") OR (#"8层下行呼梯按钮指示灯" AND (#当前楼层数 = 7) AND #"1号梯外呼上面无目标8") OR (#"9层下行呼梯按钮指示灯" AND (#当前楼层数 = 8) AND #"1号梯外呼上面无目标9")) AND #"1号梯上行接触器";
   #中间变量4 := #"1号梯下行指示" AND ((#"2层上行呼梯按钮指示灯" AND (#当前楼层数 = 3) AND #"1号梯外呼下面无目标2") OR (#"3层上行呼梯按钮指示灯" AND (#当前楼层数 = 4) AND #"1号梯外呼下面无目标3") OR (#"4层上行呼梯按钮指示灯" AND (#当前楼层数 = 5) AND #"1号梯外呼下面无目标4") OR (#"5层上行呼梯按钮指示灯" AND (#当前楼层数 = 6) AND #"1号梯外呼下面无目标5") OR (#"6层上行呼梯按钮指示灯" AND (#当前楼层数 = 7) AND #"1号梯外呼下面无目标6") OR (#"7层上行呼梯按钮指示灯" AND (#当前楼层数 = 8) AND #"1号梯外呼下面无目标7") OR (#"8层上行呼梯按钮指示灯" AND (#当前楼层数 = 9) AND #"1号梯外呼下面无目标8") OR (#"9层上行呼梯按钮指示灯" AND (#当前楼层数 = 10) AND #"1号梯外呼下面无目标9")) AND #"1号梯下行接触器";
   #将要停梯 := (#中间变量1 OR #中间变量2 OR #中间变量3 OR #中间变量4) AND NOT #"1号梯检修信号";
END_REGION

REGION Network 2: 初始化低速
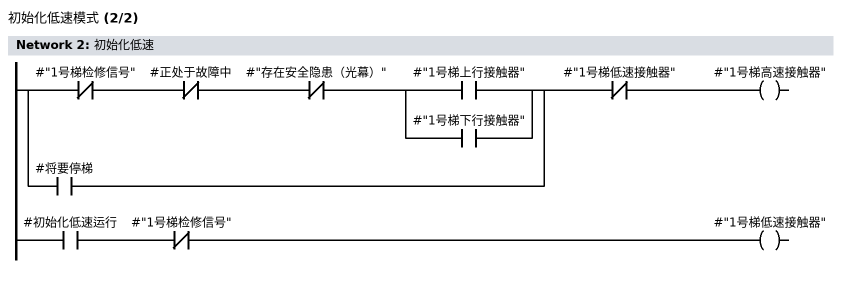
   RUNG wire#powerrail
      I_Contact( #"1号梯检修信号" )
      I_Contact( #正处于故障中 )
      I_Contact( #"存在安全隐患（光幕）" )
      wire#w1
      Contact( #"1号梯上行接触器" )
      wire#w2
      I_Contact( #"1号梯低速接触器" )
      Coil( #"1号梯高速接触器" )
   END_RUNG
   RUNG wire#w1
      Contact( #"1号梯下行接触器" )
   END_RUNG wire#w2
   RUNG wire#powerrail
      Contact( #将要停梯 )
   END_RUNG wire#w2
   RUNG wire#powerrail
      Contact( #初始化低速运行 )
      I_Contact( #"1号梯检修信号" )
      Coil( #"1号梯低速接触器" )
   END_RUNG
   // the same network as SCL:
   #"1号梯高速接触器" := ((NOT #"1号梯检修信号" AND NOT #正处于故障中 AND NOT #"存在安全隐患（光幕）" AND (#"1号梯上行接触器" OR #"1号梯下行接触器")) OR #将要停梯) AND NOT #"1号梯低速接触器";
   #"1号梯低速接触器" := #初始化低速运行 AND NOT #"1号梯检修信号";
END_REGION
END_FUNCTION_BLOCK

FUNCTION_BLOCK "上下行和制动"   // FB5, LAD
{ S7_Optimized_Access := 'TRUE' }
VERSION : 0.1
   VAR_INPUT
      载重量 : Int;
      正处于故障中 : Bool;
      "存在安全隐患（光幕）" : Bool;
      正确楼层数 : Int;
      将要停梯 : Bool;
      上平层信号 : Bool;
      下平层信号 : Bool;
      初始化将要停梯 : Bool;
      "1层上呼分配" : Bool;
      "2层上呼分配" : Bool;
      "3层上呼分配" : Bool;
      "4层上呼分配" : Bool;
      "5层上呼分配" : Bool;
      "6层上呼分配" : Bool;
      "7层上呼分配" : Bool;
      "8层上呼分配" : Bool;
      "9层上呼分配" : Bool;
      "2层下呼分配" : Bool;
      "3层下呼分配" : Bool;
      "4层下呼分配" : Bool;
      "5层下呼分配" : Bool;
      "6层下呼分配" : Bool;
      "7层下呼分配" : Bool;
      "8层下呼分配" : Bool;
      "9层下呼分配" : Bool;
      "10层下呼分配" : Bool;
      当前楼层数 : Int;
      上行指示 : Bool;
      下行指示 : Bool;
      初始化上行接触器 : Bool;
      初始化下行接触器 : Bool;
      "停梯截断(完成关门）" : Bool;
      "停梯截断(完成开门）" : Bool;
      "1号梯检修信号" : Bool;
      准备就绪 : Bool;
      "1号梯上平层信号" : Bool;
      "1号梯下平层信号" : Bool;
      "1层上行呼梯按钮" : Bool;
      "2层上行呼梯按钮" : Bool;
      "3层上行呼梯按钮" : Bool;
      "4层上行呼梯按钮" : Bool;
      "5层上行呼梯按钮" : Bool;
      "6层上行呼梯按钮" : Bool;
      "7层上行呼梯按钮" : Bool;
      "8层上行呼梯按钮" : Bool;
      "9层上行呼梯按钮" : Bool;
      "2层下行呼梯按钮" : Bool;
      "3层下行呼梯按钮" : Bool;
      "4层下行呼梯按钮" : Bool;
      "5层下行呼梯按钮" : Bool;
      "6层下行呼梯按钮" : Bool;
      "7层下行呼梯按钮" : Bool;
      "8层下行呼梯按钮" : Bool;
      "9层下行呼梯按钮" : Bool;
      "10层下行呼梯按钮" : Bool;
      "1号梯轿内选层按钮1" : Bool;
      "1号梯轿内选层按钮2" : Bool;
      "1号梯轿内选层按钮3" : Bool;
      "1号梯轿内选层按钮4" : Bool;
      "1号梯轿内选层按钮5" : Bool;
      "1号梯轿内选层按钮6" : Bool;
      "1号梯轿内选层按钮7" : Bool;
      "1号梯轿内选层按钮8" : Bool;
      "1号梯轿内选层按钮9" : Bool;
      "1号梯轿内选层按钮10" : Bool;
      死机 : Bool;
      满载指示 : Bool;
   END_VAR
   VAR_OUTPUT
      就近运动电梯 : Bool;
      "1号梯上行指示" : Bool;
      "1号梯下行指示" : Bool;
      上行接触器 : Bool;
      下行接触器 : Bool;
      "1号梯1层按钮指示灯" : Bool;
      "1号梯2层按钮指示灯" : Bool;
      "1号梯3层按钮指示灯" : Bool;
      "1号梯4层按钮指示灯" : Bool;
      "1号梯5层按钮指示灯" : Bool;
      "1号梯6层按钮指示灯" : Bool;
      "1号梯7层按钮指示灯" : Bool;
      "1号梯8层按钮指示灯" : Bool;
      "1号梯9层按钮指示灯" : Bool;
      "1号梯10层按钮指示灯" : Bool;
      "1号梯1级减速制动" : Bool;
      "1号梯2级减速制动" : Bool;
      "1号梯3级减速制动" : Bool;
   END_VAR
   VAR
      中间关断 : Bool;
      梯内有人不走 : Bool;
      刚刚在上行 : Bool;
      刚刚在下行 : Bool;
      准备刹车 : Bool;
      连接1 : Bool;
      优先停梯1 : Bool;
      优先停梯2 : Bool;
      客人有下行需求后延迟下行指示a : TOF_TIME;
      客人有上行需求后延迟上行指示a : TOF_TIME;
      IEC_Timer_0_Instance : TON_TIME;
      卡顿上行 : Bool;
      卡顿下行 : Bool;
      卡顿制速 : Bool;
      连接11 : Bool;
      连接13 : Bool;
      连接14 : Bool;
      连接15 : Bool;
      连接16 : Bool;
      连接18 : Bool;
      连接19 : Bool;
      连接20 : Bool;
      连接21 : Bool;
      连接23 : Bool;
      连接24 : Bool;
      连接25 : Bool;
      连接26 : Bool;
      连接28 : Bool;
      连接29 : Bool;
      连接30 : Bool;
      连接31 : Bool;
      连接33 : Bool;
      连接34 : Bool;
      连接35 : Bool;
      连接36 : Bool;
      连接37 : Bool;
      连接38 : Bool;
      连接39 : Bool;
      连接40 : Bool;
      连接41 : Bool;
      连接42 : Bool;
      连接43 : Bool;
      连接44 : Bool;
      连接45 : Bool;
      连接46 : Bool;
      连接47 : Bool;
      连接74 : Bool;
      连接75 : Bool;
      连接76 : Bool;
      连接77 : Bool;
      连接78 : Bool;
      连接79 : Bool;
      连接80 : Bool;
      连接81 : Bool;
      连接82 : Bool;
      连接83 : Bool;
      连接84 : Bool;
      连接85 : Bool;
      连接86 : Bool;
      连接87 : Bool;
      连接88 : Bool;
      连接89 : Bool;
      连接90 : Bool;
      连接91 : Bool;
      连接92 : Bool;
      连接93 : Bool;
      连接94 : Bool;
      连接95 : Bool;
      连接96 : Bool;
      连接97 : Bool;
      连接98 : Bool;
      连接99 : Bool;
      连接100 : Bool;
      连接102 : Bool;
      连接103 : Bool;
      连接104 : Bool;
      连接105 : Bool;
      电梯停止后延时灭灯2楼上 : TON_TIME;
      电梯停止后延时灭灯3楼上 : TON_TIME;
      电梯停止后延时灭灯4楼上 : TON_TIME;
      电梯停止后延时灭灯5楼上 : TON_TIME;
      电梯停止后延时灭灯6楼上 : TON_TIME;
      电梯停止后延时灭灯7楼上 : TON_TIME;
      电梯停止后延时灭灯8楼上 : TON_TIME;
      电梯停止后延时灭灯9楼上 : TON_TIME;
      电梯停止后延时灭灯2楼下 : TON_TIME;
      电梯停止后延时灭灯3楼下 : TON_TIME;
      电梯停止后延时灭灯4楼下 : TON_TIME;
      停止后延时灭灯5楼下 : TON_TIME;
      电梯停止后延时灭灯6楼下 : TON_TIME;
      电梯停止后延时灭灯7楼下 : TON_TIME;
      电梯停止后延时灭灯8楼下 : TON_TIME;
      电梯停止后延时灭灯9楼下 : TON_TIME;
      "电梯停止后延时灭灯 1楼" : TON_TIME;
      "电梯停止后延时灭灯 10楼" : TON_TIME;
      连接2 : Bool;
      IEC_Timer_0_Instance_1 : TOF_TIME;
      IEC_Timer_0_Instance_2 : TON_TIME;
      IEC_Timer_0_Instance_3 : TOF_TIME;
      IEC_Timer_0_Instance_7 : TOF_TIME;
      "IEC _Timer_0_Instance_6" : TON_TIME;
      IEC_Timer_0_Instance_4 : TON_TIME;
      IEC_Timr_0_Instance_5 : TP_TIME;
   END_VAR
   VAR RETAIN
      IEC_Counter_0_Instance : CTU_INT;
   END_VAR
   VAR
      满载关灯 : Bool;
      IEC_Timer_0_Instance_5 : TON_TIME;
   END_VAR
   VAR RETAIN
      IEC_Counter_0_Instance_1 : CTU_INT;
   END_VAR
   VAR
      中间1 : Bool;
      IEC_Timer_0_Instance_6 : TP_TIME;
   END_VAR
   VAR_TEMP   // added for the SCL form of the ladder/FBD networks
      _w1 : Bool;
      _w2 : Bool;
      _w3 : Bool;
      _w4 : Bool;
      _w5 : Bool;
      _w6 : Bool;
      _w7 : Bool;
      _w8 : Bool;
      _w9 : Bool;
      _w10 : Bool;
      _w11 : Bool;
      _w12 : Bool;
      _w13 : Bool;
      _w14 : Bool;
      _w15 : Bool;
      _w16 : Bool;
      _w17 : Bool;
      _w18 : Bool;
      _w19 : Bool;
      _w20 : Bool;
      _w21 : Bool;
      _w22 : Bool;
      _w23 : Bool;
      _w24 : Bool;
      _w25 : Bool;
      _w26 : Bool;
      _w27 : Bool;
      _w28 : Bool;
      _w29 : Bool;
      _w30 : Bool;
      _w31 : Bool;
      _w32 : Bool;
   END_VAR
BEGIN

REGION Network 1: 上下行接触器
   // 用“停梯优先级”里的‘停梯截断’优先控制 停 ，再用“开关门”里的‘完成开门关门’严格控制 动
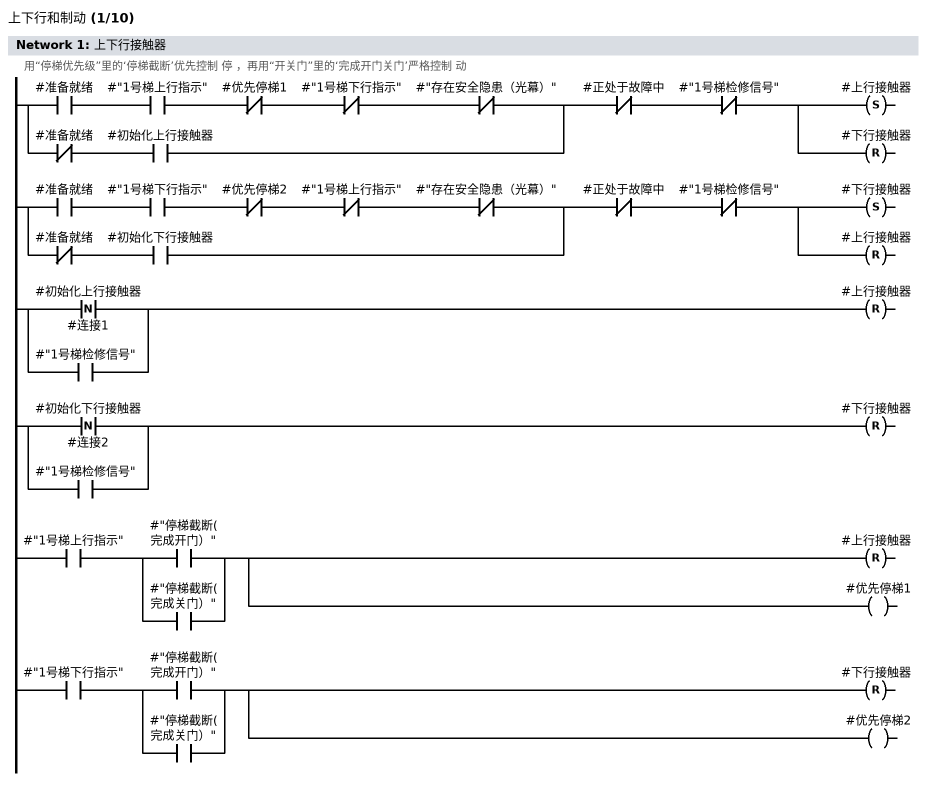
   RUNG wire#powerrail
      Contact( #准备就绪 )
      Contact( #"1号梯上行指示" )
      I_Contact( #优先停梯1 )
      I_Contact( #"1号梯下行指示" )
      I_Contact( #"存在安全隐患（光幕）" )
      wire#w1
      I_Contact( #正处于故障中 )
      I_Contact( #"1号梯检修信号" )
      wire#w2
      S_Coil( #上行接触器 )
   END_RUNG
   RUNG wire#powerrail
      I_Contact( #准备就绪 )
      Contact( #初始化上行接触器 )
   END_RUNG wire#w1
   RUNG wire#w2
      R_Coil( #下行接触器 )
   END_RUNG
   RUNG wire#powerrail
      Contact( #准备就绪 )
      Contact( #"1号梯下行指示" )
      I_Contact( #优先停梯2 )
      I_Contact( #"1号梯上行指示" )
      I_Contact( #"存在安全隐患（光幕）" )
      wire#w3
      I_Contact( #正处于故障中 )
      I_Contact( #"1号梯检修信号" )
      wire#w4
      S_Coil( #下行接触器 )
   END_RUNG
   RUNG wire#powerrail
      I_Contact( #准备就绪 )
      Contact( #初始化下行接触器 )
   END_RUNG wire#w3
   RUNG wire#w4
      R_Coil( #上行接触器 )
   END_RUNG
   RUNG wire#powerrail
      N_Contact(operand := #初始化上行接触器, bit := #连接1)
      wire#w5
      R_Coil( #上行接触器 )
   END_RUNG
   RUNG wire#powerrail
      Contact( #"1号梯检修信号" )
   END_RUNG wire#w5
   RUNG wire#powerrail
      N_Contact(operand := #初始化下行接触器, bit := #连接2)
      wire#w6
      R_Coil( #下行接触器 )
   END_RUNG
   RUNG wire#powerrail
      Contact( #"1号梯检修信号" )
   END_RUNG wire#w6
   RUNG wire#powerrail
      Contact( #"1号梯上行指示" )
      wire#w7
      Contact( #"停梯截断(完成开门）" )
      wire#w8
      R_Coil( #上行接触器 )
   END_RUNG
   RUNG wire#w7
      Contact( #"停梯截断(完成关门）" )
   END_RUNG wire#w8
   RUNG wire#w8
      Coil( #优先停梯1 )
   END_RUNG
   RUNG wire#powerrail
      Contact( #"1号梯下行指示" )
      wire#w9
      Contact( #"停梯截断(完成开门）" )
      wire#w10
      R_Coil( #下行接触器 )
   END_RUNG
   RUNG wire#w9
      Contact( #"停梯截断(完成关门）" )
   END_RUNG wire#w10
   RUNG wire#w10
      Coil( #优先停梯2 )
   END_RUNG
   // the same network as SCL:
   IF ((#准备就绪 AND #"1号梯上行指示" AND NOT #优先停梯1 AND NOT #"1号梯下行指示" AND NOT #"存在安全隐患（光幕）") OR (NOT #准备就绪 AND #初始化上行接触器)) AND NOT #正处于故障中 AND NOT #"1号梯检修信号" THEN
       #上行接触器 := TRUE;
       #下行接触器 := FALSE;
   END_IF;
   IF ((#准备就绪 AND #"1号梯下行指示" AND NOT #优先停梯2 AND NOT #"1号梯上行指示" AND NOT #"存在安全隐患（光幕）") OR (NOT #准备就绪 AND #初始化下行接触器)) AND NOT #正处于故障中 AND NOT #"1号梯检修信号" THEN
       #下行接触器 := TRUE;
       #上行接触器 := FALSE;
   END_IF;
   #_w1 := NOT #初始化上行接触器 AND #连接1;   // falling edge of #初始化上行接触器
   #连接1 := #初始化上行接触器;
   IF #_w1 OR #"1号梯检修信号" THEN #上行接触器 := FALSE; END_IF;
   #_w2 := NOT #初始化下行接触器 AND #连接2;   // falling edge of #初始化下行接触器
   #连接2 := #初始化下行接触器;
   IF #_w2 OR #"1号梯检修信号" THEN #下行接触器 := FALSE; END_IF;
   #_w3 := #"1号梯上行指示" AND (#"停梯截断(完成开门）" OR #"停梯截断(完成关门）");
   IF #_w3 THEN #上行接触器 := FALSE; END_IF;
   #优先停梯1 := #_w3;
   #_w4 := #"1号梯下行指示" AND (#"停梯截断(完成开门）" OR #"停梯截断(完成关门）");
   IF #_w4 THEN #下行接触器 := FALSE; END_IF;
   #优先停梯2 := #_w4;
END_REGION

REGION Network 2: 应对卡顿的 继续上下行指示
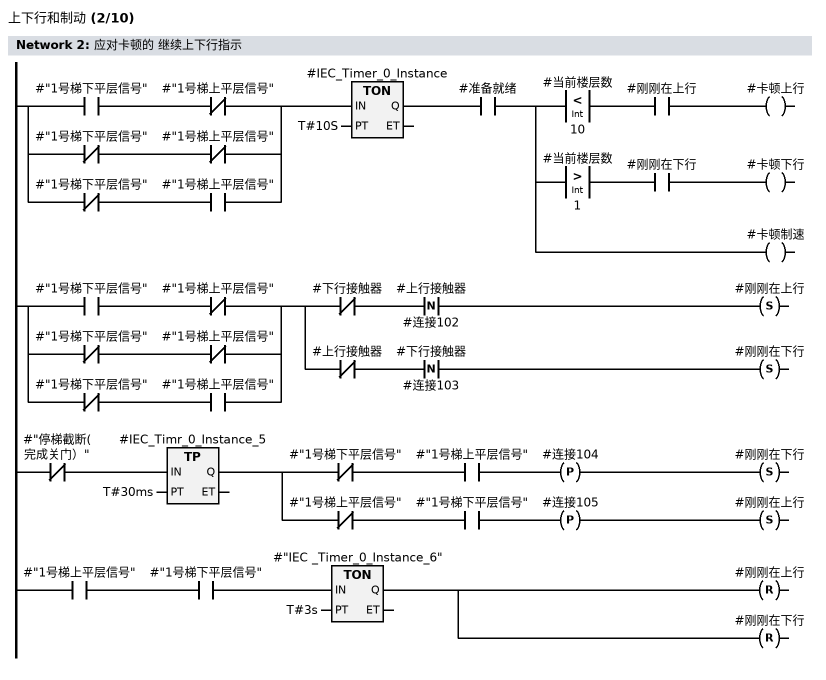
   #IEC_Timer_0_Instance(IN := (#"1号梯下平层信号" AND NOT #"1号梯上平层信号") OR (NOT #"1号梯下平层信号" AND NOT #"1号梯上平层信号") OR (NOT #"1号梯下平层信号" AND #"1号梯上平层信号"),   // TON
                         PT := T#10S);
   #_w1 := #IEC_Timer_0_Instance.Q AND #准备就绪;
   #卡顿上行 := #_w1 AND (#当前楼层数 < 10) AND #刚刚在上行;
   #卡顿下行 := #_w1 AND (#当前楼层数 > 1) AND #刚刚在下行;
   #卡顿制速 := #_w1;
   #_w2 := (#"1号梯下平层信号" AND NOT #"1号梯上平层信号") OR (NOT #"1号梯下平层信号" AND NOT #"1号梯上平层信号") OR (NOT #"1号梯下平层信号" AND #"1号梯上平层信号");
   #_w3 := #_w2 AND NOT #下行接触器 AND NOT #上行接触器 AND #连接102;   // falling edge of #上行接触器
   #连接102 := #上行接触器;
   IF #_w3 THEN #刚刚在上行 := TRUE; END_IF;
   #_w4 := #_w2 AND NOT #上行接触器 AND NOT #下行接触器 AND #连接103;   // falling edge of #下行接触器
   #连接103 := #下行接触器;
   IF #_w4 THEN #刚刚在下行 := TRUE; END_IF;
   #IEC_Timr_0_Instance_5(IN := NOT #"停梯截断(完成关门）", PT := T#30ms);   // TP
   #_w5 := #IEC_Timr_0_Instance_5.Q AND NOT #"1号梯下平层信号" AND #"1号梯上平层信号";
   #_w6 := #_w5 AND NOT #连接104;   // rising edge
   #连接104 := #_w5;
   IF #_w6 THEN #刚刚在下行 := TRUE; END_IF;
   #_w7 := #IEC_Timr_0_Instance_5.Q AND NOT #"1号梯上平层信号" AND #"1号梯下平层信号";
   #_w8 := #_w7 AND NOT #连接105;   // rising edge
   #连接105 := #_w7;
   IF #_w8 THEN #刚刚在上行 := TRUE; END_IF;
   #"IEC _Timer_0_Instance_6"(IN := #"1号梯上平层信号" AND #"1号梯下平层信号", PT := T#3s);   // TON
   IF #"IEC _Timer_0_Instance_6".Q THEN
       #刚刚在上行 := FALSE;
       #刚刚在下行 := FALSE;
   END_IF;
END_REGION

REGION Network 3: 上行指示
   // （不考虑先后级）
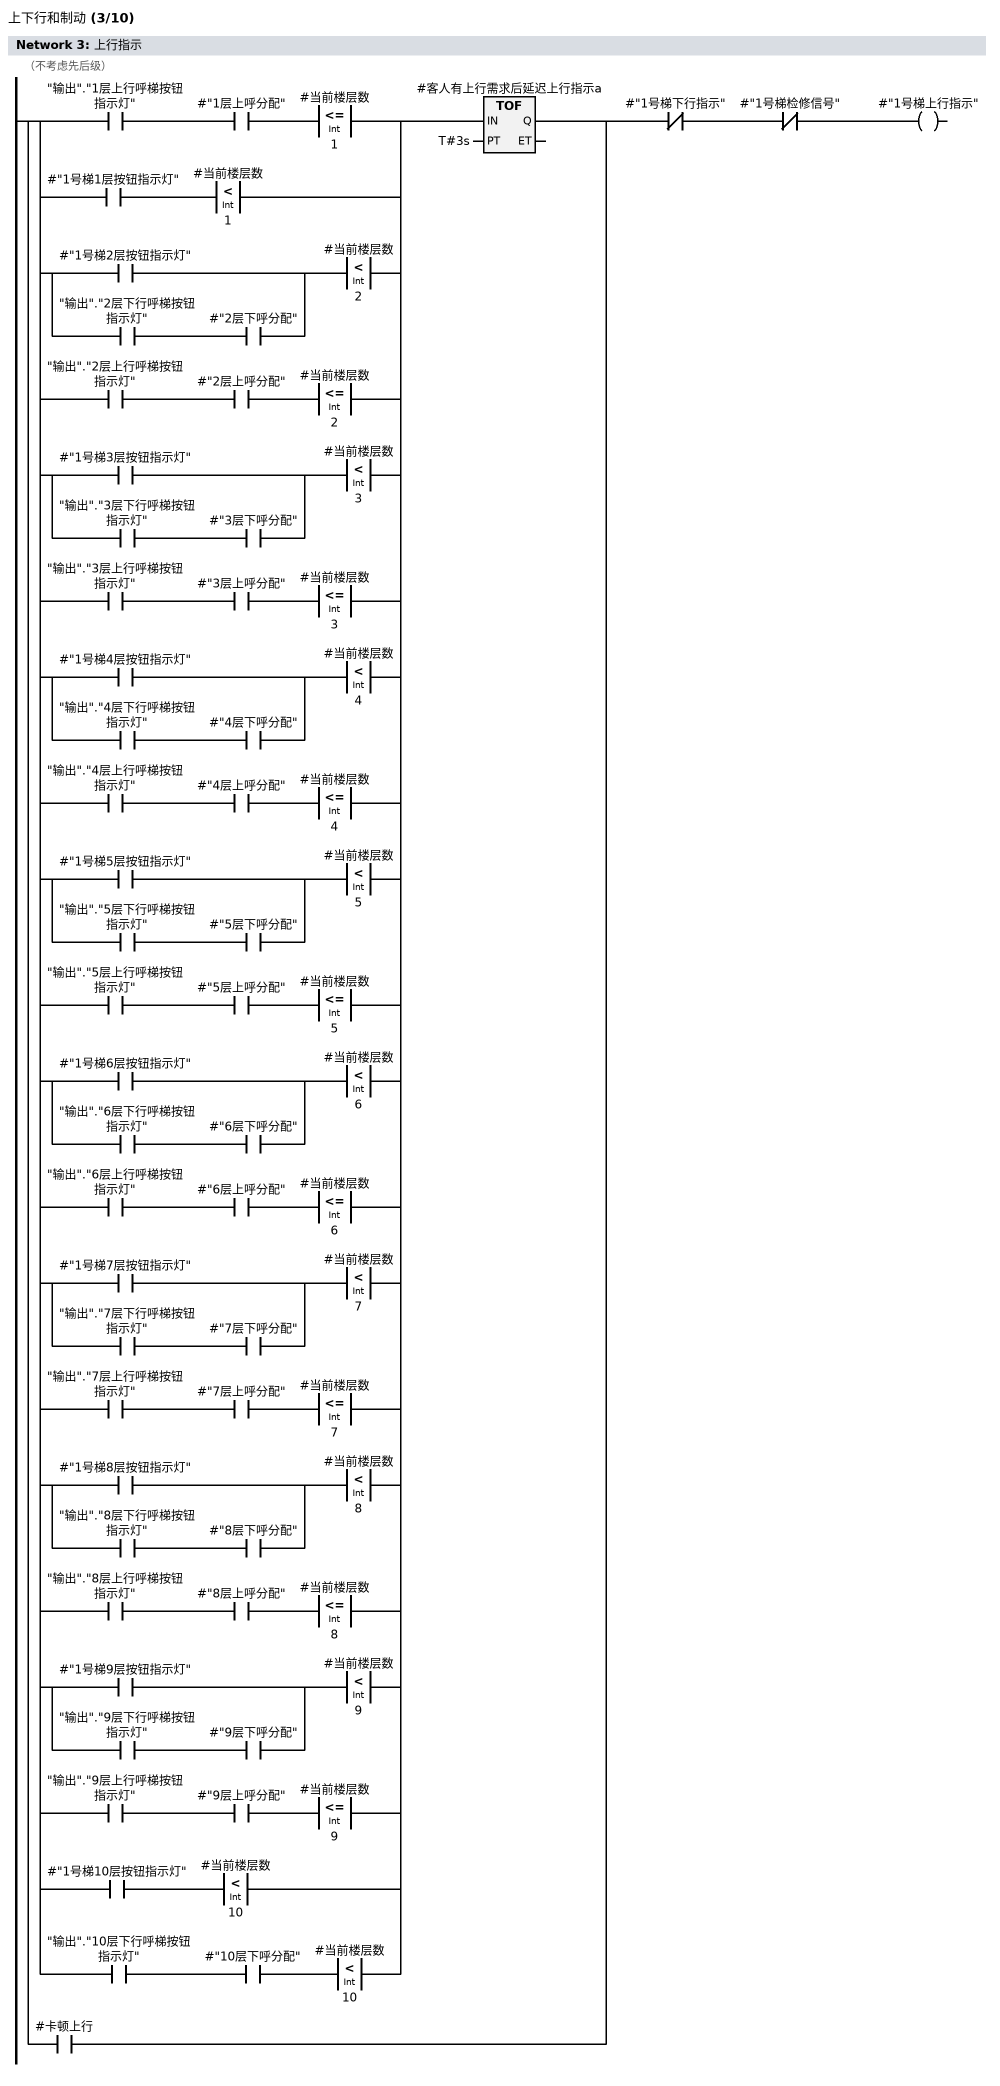
   #客人有上行需求后延迟上行指示a(IN := ("输出"."1层上行呼梯按钮指示灯" AND #"1层上呼分配" AND (#当前楼层数 <= 1)) OR (#"1号梯1层按钮指示灯" AND (#当前楼层数 < 1)) OR ((#"1号梯2层按钮指示灯" OR ("输出"."2层下行呼梯按钮指示灯" AND #"2层下呼分配")) AND (#当前楼层数 < 2)) OR ("输出"."2层上行呼梯按钮指示灯" AND #"2层上呼分配" AND (#当前楼层数 <= 2)) OR ((#"1号梯3层按钮指示灯" OR ("输出"."3层下行呼梯按钮指示灯" AND #"3层下呼分配")) AND (#当前楼层数 < 3)) OR ("输出"."3层上行呼梯按钮指示灯" AND #"3层上呼分配" AND (#当前楼层数 <= 3)) OR ((#"1号梯4层按钮指示灯" OR ("输出"."4层下行呼梯按钮指示灯" AND #"4层下呼分配")) AND (#当前楼层数 < 4)) OR ("输出"."4层上行呼梯按钮指示灯" AND #"4层上呼分配" AND (#当前楼层数 <= 4)) OR ((#"1号梯5层按钮指示灯" OR ("输出"."5层下行呼梯按钮指示灯" AND #"5层下呼分配")) AND (#当前楼层数 < 5)) OR ("输出"."5层上行呼梯按钮指示灯" AND #"5层上呼分配" AND (#当前楼层数 <= 5)) OR ((#"1号梯6层按钮指示灯" OR ("输出"."6层下行呼梯按钮指示灯" AND #"6层下呼分配")) AND (#当前楼层数 < 6)) OR ("输出"."6层上行呼梯按钮指示灯" AND #"6层上呼分配" AND (#当前楼层数 <= 6)) OR ((#"1号梯7层按钮指示灯" OR ("输出"."7层下行呼梯按钮指示灯" AND #"7层下呼分配")) AND (#当前楼层数 < 7)) OR ("输出"."7层上行呼梯按钮指示灯" AND #"7层上呼分配" AND (#当前楼层数 <= 7)) OR ((#"1号梯8层按钮指示灯" OR ("输出"."8层下行呼梯按钮指示灯" AND #"8层下呼分配")) AND (#当前楼层数 < 8)) OR ("输出"."8层上行呼梯按钮指示灯" AND #"8层上呼分配" AND (#当前楼层数 <= 8)) OR ((#"1号梯9层按钮指示灯" OR ("输出"."9层下行呼梯按钮指示灯" AND #"9层下呼分配")) AND (#当前楼层数 < 9)) OR ("输出"."9层上行呼梯按钮指示灯" AND #"9层上呼分配" AND (#当前楼层数 <= 9)) OR (#"1号梯10层按钮指示灯" AND (#当前楼层数 < 10)) OR ("输出"."10层下行呼梯按钮指示灯" AND #"10层下呼分配" AND (#当前楼层数 < 10)),   // TOF
                    PT := T#3s);
   #"1号梯上行指示" := (#客人有上行需求后延迟上行指示a.Q OR #卡顿上行) AND NOT #"1号梯下行指示" AND NOT #"1号梯检修信号";
END_REGION

REGION Network 4: 下行指示
   // （不考虑优先级）
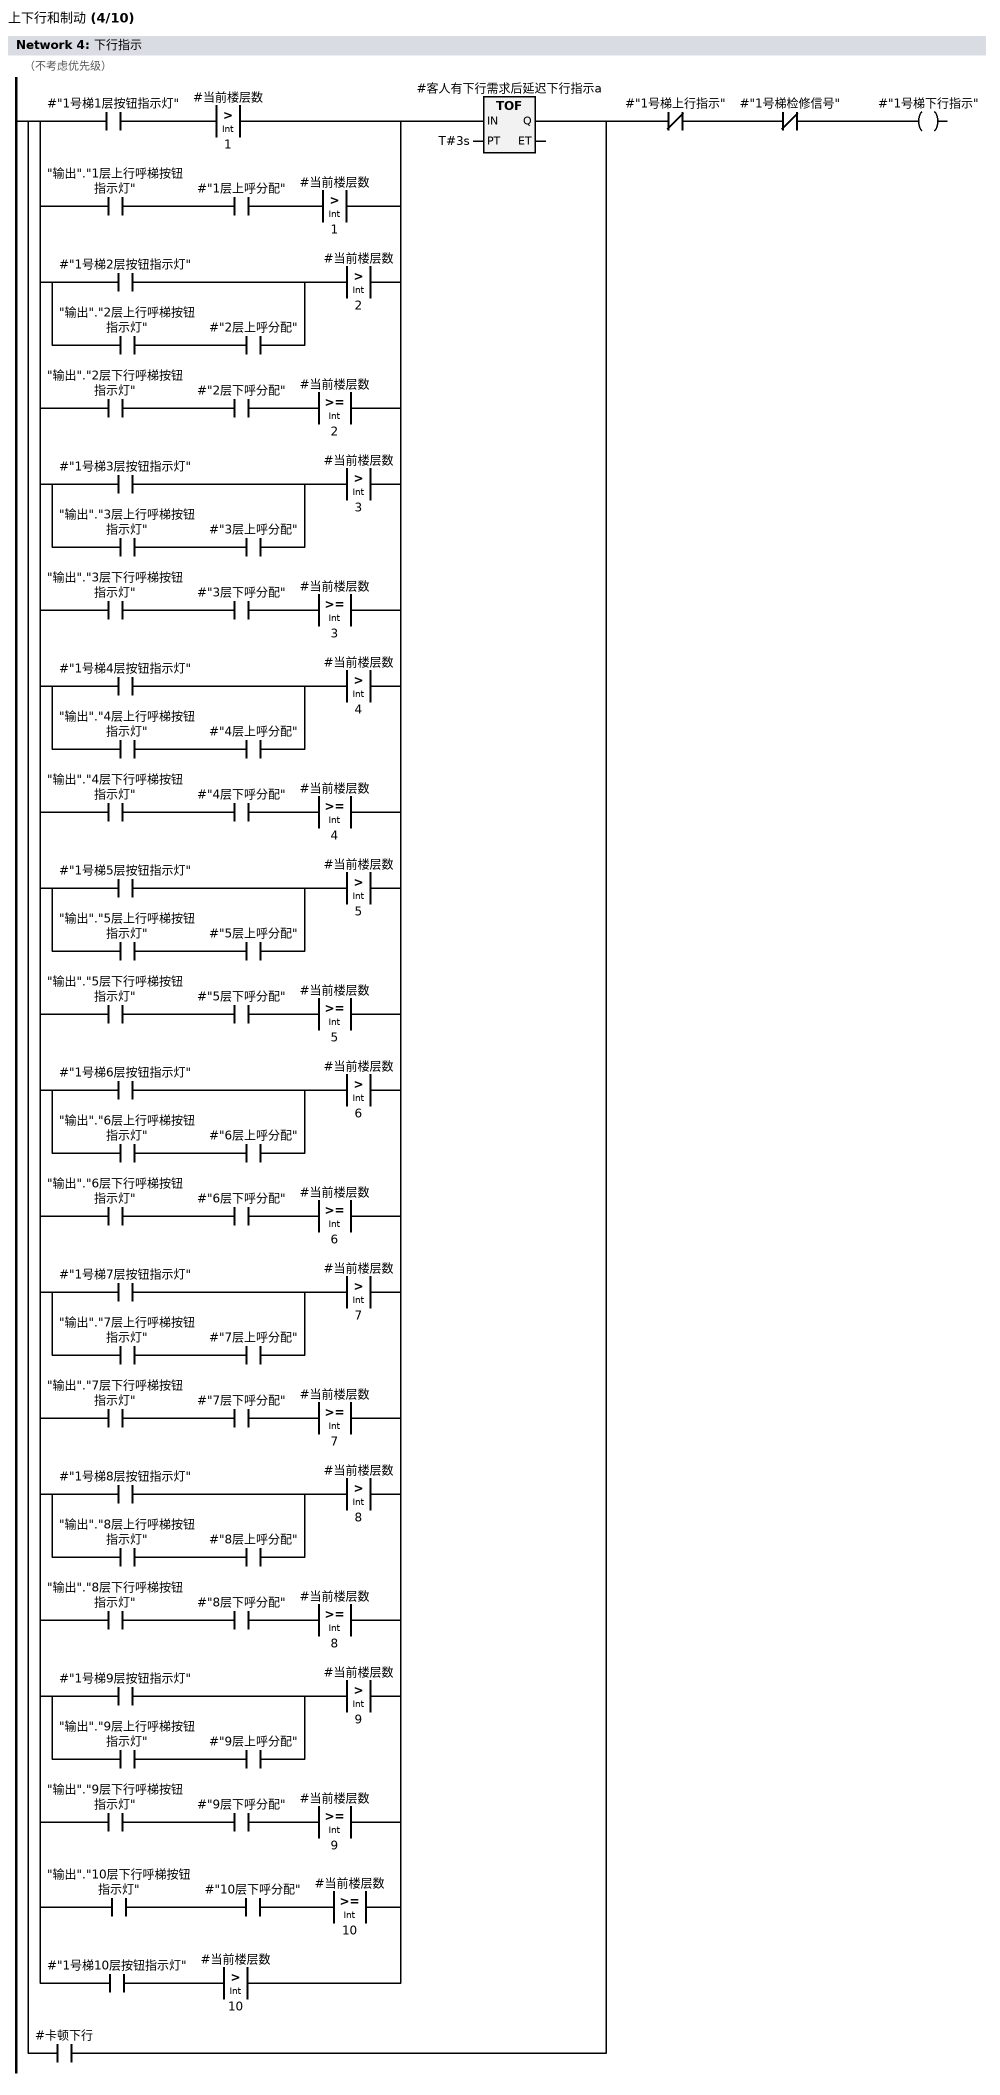
   #客人有下行需求后延迟下行指示a(IN := (#"1号梯1层按钮指示灯" AND (#当前楼层数 > 1)) OR ("输出"."1层上行呼梯按钮指示灯" AND #"1层上呼分配" AND (#当前楼层数 > 1)) OR ((#"1号梯2层按钮指示灯" OR ("输出"."2层上行呼梯按钮指示灯" AND #"2层上呼分配")) AND (#当前楼层数 > 2)) OR ("输出"."2层下行呼梯按钮指示灯" AND #"2层下呼分配" AND (#当前楼层数 >= 2)) OR ((#"1号梯3层按钮指示灯" OR ("输出"."3层上行呼梯按钮指示灯" AND #"3层上呼分配")) AND (#当前楼层数 > 3)) OR ("输出"."3层下行呼梯按钮指示灯" AND #"3层下呼分配" AND (#当前楼层数 >= 3)) OR ((#"1号梯4层按钮指示灯" OR ("输出"."4层上行呼梯按钮指示灯" AND #"4层上呼分配")) AND (#当前楼层数 > 4)) OR ("输出"."4层下行呼梯按钮指示灯" AND #"4层下呼分配" AND (#当前楼层数 >= 4)) OR ((#"1号梯5层按钮指示灯" OR ("输出"."5层上行呼梯按钮指示灯" AND #"5层上呼分配")) AND (#当前楼层数 > 5)) OR ("输出"."5层下行呼梯按钮指示灯" AND #"5层下呼分配" AND (#当前楼层数 >= 5)) OR ((#"1号梯6层按钮指示灯" OR ("输出"."6层上行呼梯按钮指示灯" AND #"6层上呼分配")) AND (#当前楼层数 > 6)) OR ("输出"."6层下行呼梯按钮指示灯" AND #"6层下呼分配" AND (#当前楼层数 >= 6)) OR ((#"1号梯7层按钮指示灯" OR ("输出"."7层上行呼梯按钮指示灯" AND #"7层上呼分配")) AND (#当前楼层数 > 7)) OR ("输出"."7层下行呼梯按钮指示灯" AND #"7层下呼分配" AND (#当前楼层数 >= 7)) OR ((#"1号梯8层按钮指示灯" OR ("输出"."8层上行呼梯按钮指示灯" AND #"8层上呼分配")) AND (#当前楼层数 > 8)) OR ("输出"."8层下行呼梯按钮指示灯" AND #"8层下呼分配" AND (#当前楼层数 >= 8)) OR ((#"1号梯9层按钮指示灯" OR ("输出"."9层上行呼梯按钮指示灯" AND #"9层上呼分配")) AND (#当前楼层数 > 9)) OR ("输出"."9层下行呼梯按钮指示灯" AND #"9层下呼分配" AND (#当前楼层数 >= 9)) OR ("输出"."10层下行呼梯按钮指示灯" AND #"10层下呼分配" AND (#当前楼层数 >= 10)) OR (#"1号梯10层按钮指示灯" AND (#当前楼层数 > 10)),   // TOF
                    PT := T#3s);
   #"1号梯下行指示" := (#客人有下行需求后延迟下行指示a.Q OR #卡顿下行) AND NOT #"1号梯上行指示" AND NOT #"1号梯检修信号";
END_REGION

REGION Network 5: 1楼和10楼 的外呼按钮和指示灯
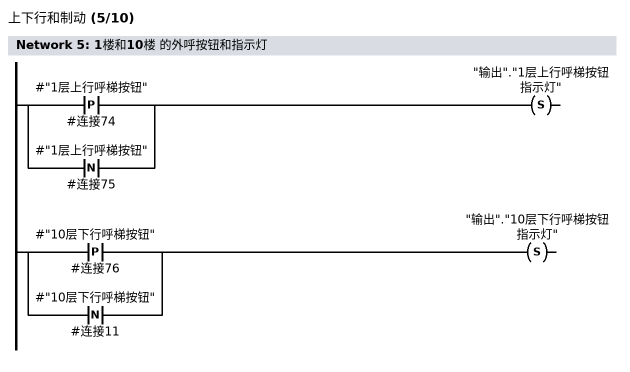
   RUNG wire#powerrail
      P_Contact(operand := #"1层上行呼梯按钮", bit := #连接74)
      wire#w1
      S_Coil( "输出"."1层上行呼梯按钮指示灯" )
   END_RUNG
   RUNG wire#powerrail
      N_Contact(operand := #"1层上行呼梯按钮", bit := #连接75)
   END_RUNG wire#w1
   RUNG wire#powerrail
      P_Contact(operand := #"10层下行呼梯按钮", bit := #连接76)
      wire#w2
      S_Coil( "输出"."10层下行呼梯按钮指示灯" )
   END_RUNG
   RUNG wire#powerrail
      N_Contact(operand := #"10层下行呼梯按钮", bit := #连接11)
   END_RUNG wire#w2
   // the same network as SCL:
   #_w1 := #"1层上行呼梯按钮" AND NOT #连接74;   // rising edge of #"1层上行呼梯按钮"
   #连接74 := #"1层上行呼梯按钮";
   #_w2 := NOT #"1层上行呼梯按钮" AND #连接75;   // falling edge of #"1层上行呼梯按钮"
   #连接75 := #"1层上行呼梯按钮";
   IF #_w1 OR #_w2 THEN "输出"."1层上行呼梯按钮指示灯" := TRUE; END_IF;
   #_w3 := #"10层下行呼梯按钮" AND NOT #连接76;   // rising edge of #"10层下行呼梯按钮"
   #连接76 := #"10层下行呼梯按钮";
   #_w4 := NOT #"10层下行呼梯按钮" AND #连接11;   // falling edge of #"10层下行呼梯按钮"
   #连接11 := #"10层下行呼梯按钮";
   IF #_w3 OR #_w4 THEN "输出"."10层下行呼梯按钮指示灯" := TRUE; END_IF;
END_REGION

REGION Network 6: 2~4楼外呼 按钮和指示灯
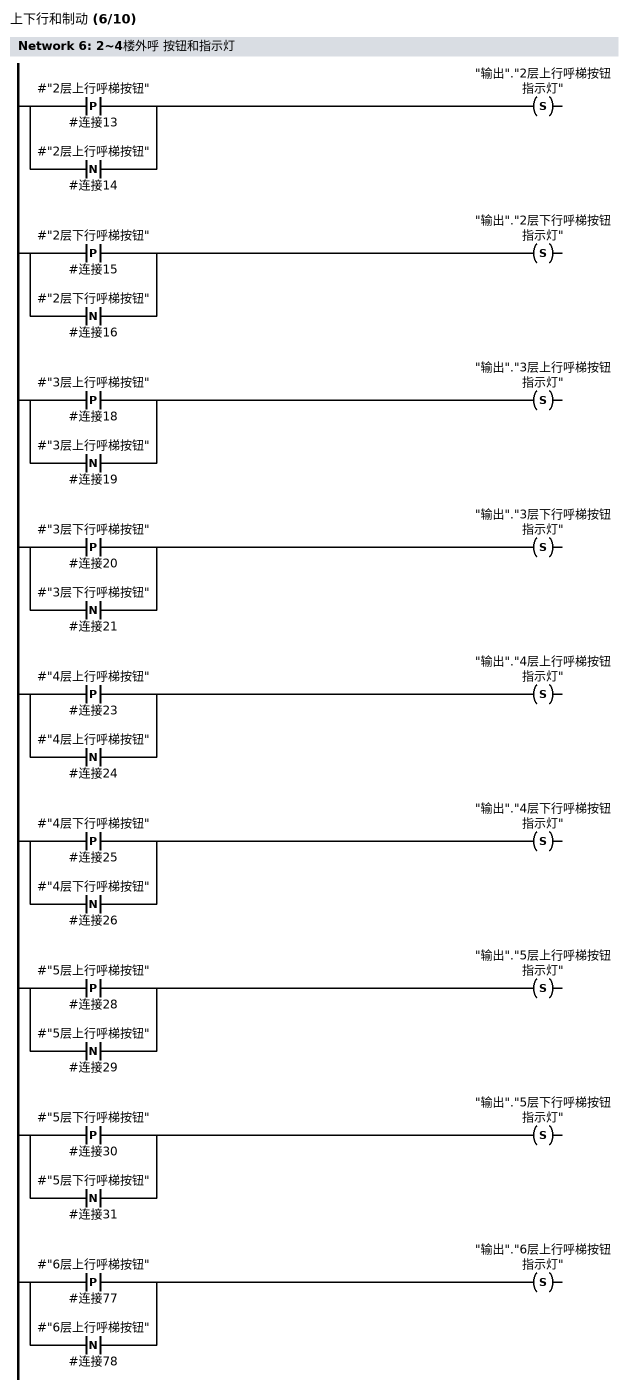
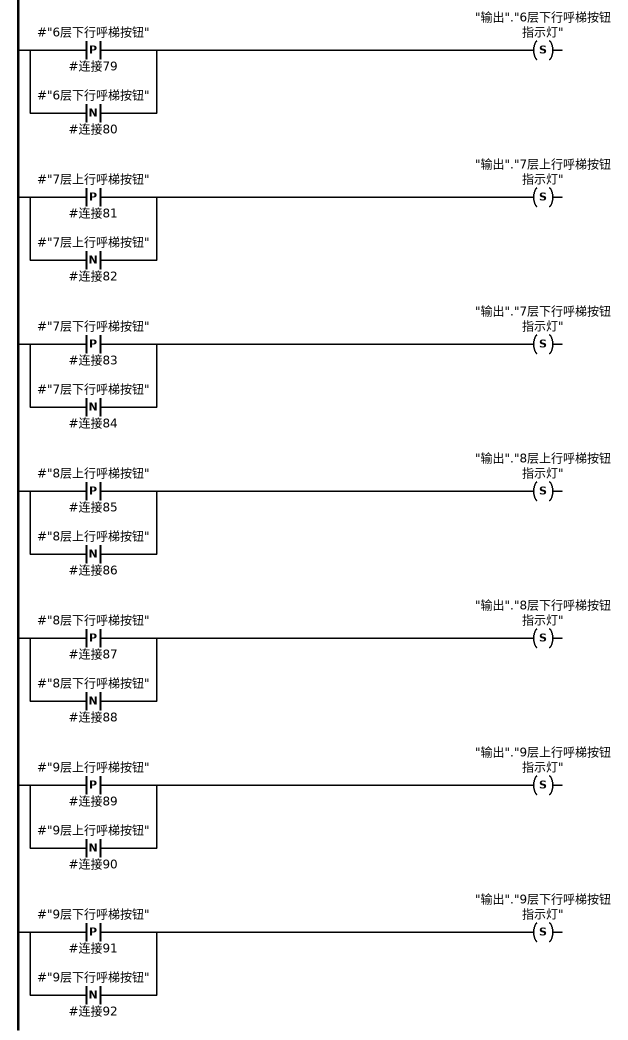
   RUNG wire#powerrail
      P_Contact(operand := #"2层上行呼梯按钮", bit := #连接13)
      wire#w1
      S_Coil( "输出"."2层上行呼梯按钮指示灯" )
   END_RUNG
   RUNG wire#powerrail
      N_Contact(operand := #"2层上行呼梯按钮", bit := #连接14)
   END_RUNG wire#w1
   RUNG wire#powerrail
      P_Contact(operand := #"2层下行呼梯按钮", bit := #连接15)
      wire#w2
      S_Coil( "输出"."2层下行呼梯按钮指示灯" )
   END_RUNG
   RUNG wire#powerrail
      N_Contact(operand := #"2层下行呼梯按钮", bit := #连接16)
   END_RUNG wire#w2
   RUNG wire#powerrail
      P_Contact(operand := #"3层上行呼梯按钮", bit := #连接18)
      wire#w3
      S_Coil( "输出"."3层上行呼梯按钮指示灯" )
   END_RUNG
   RUNG wire#powerrail
      N_Contact(operand := #"3层上行呼梯按钮", bit := #连接19)
   END_RUNG wire#w3
   RUNG wire#powerrail
      P_Contact(operand := #"3层下行呼梯按钮", bit := #连接20)
      wire#w4
      S_Coil( "输出"."3层下行呼梯按钮指示灯" )
   END_RUNG
   RUNG wire#powerrail
      N_Contact(operand := #"3层下行呼梯按钮", bit := #连接21)
   END_RUNG wire#w4
   RUNG wire#powerrail
      P_Contact(operand := #"4层上行呼梯按钮", bit := #连接23)
      wire#w5
      S_Coil( "输出"."4层上行呼梯按钮指示灯" )
   END_RUNG
   RUNG wire#powerrail
      N_Contact(operand := #"4层上行呼梯按钮", bit := #连接24)
   END_RUNG wire#w5
   RUNG wire#powerrail
      P_Contact(operand := #"4层下行呼梯按钮", bit := #连接25)
      wire#w6
      S_Coil( "输出"."4层下行呼梯按钮指示灯" )
   END_RUNG
   RUNG wire#powerrail
      N_Contact(operand := #"4层下行呼梯按钮", bit := #连接26)
   END_RUNG wire#w6
   RUNG wire#powerrail
      P_Contact(operand := #"5层上行呼梯按钮", bit := #连接28)
      wire#w7
      S_Coil( "输出"."5层上行呼梯按钮指示灯" )
   END_RUNG
   RUNG wire#powerrail
      N_Contact(operand := #"5层上行呼梯按钮", bit := #连接29)
   END_RUNG wire#w7
   RUNG wire#powerrail
      P_Contact(operand := #"5层下行呼梯按钮", bit := #连接30)
      wire#w8
      S_Coil( "输出"."5层下行呼梯按钮指示灯" )
   END_RUNG
   RUNG wire#powerrail
      N_Contact(operand := #"5层下行呼梯按钮", bit := #连接31)
   END_RUNG wire#w8
   RUNG wire#powerrail
      P_Contact(operand := #"6层上行呼梯按钮", bit := #连接77)
      wire#w9
      S_Coil( "输出"."6层上行呼梯按钮指示灯" )
   END_RUNG
   RUNG wire#powerrail
      N_Contact(operand := #"6层上行呼梯按钮", bit := #连接78)
   END_RUNG wire#w9
   RUNG wire#powerrail
      P_Contact(operand := #"6层下行呼梯按钮", bit := #连接79)
      wire#w10
      S_Coil( "输出"."6层下行呼梯按钮指示灯" )
   END_RUNG
   RUNG wire#powerrail
      N_Contact(operand := #"6层下行呼梯按钮", bit := #连接80)
   END_RUNG wire#w10
   RUNG wire#powerrail
      P_Contact(operand := #"7层上行呼梯按钮", bit := #连接81)
      wire#w11
      S_Coil( "输出"."7层上行呼梯按钮指示灯" )
   END_RUNG
   RUNG wire#powerrail
      N_Contact(operand := #"7层上行呼梯按钮", bit := #连接82)
   END_RUNG wire#w11
   RUNG wire#powerrail
      P_Contact(operand := #"7层下行呼梯按钮", bit := #连接83)
      wire#w12
      S_Coil( "输出"."7层下行呼梯按钮指示灯" )
   END_RUNG
   RUNG wire#powerrail
      N_Contact(operand := #"7层下行呼梯按钮", bit := #连接84)
   END_RUNG wire#w12
   RUNG wire#powerrail
      P_Contact(operand := #"8层上行呼梯按钮", bit := #连接85)
      wire#w13
      S_Coil( "输出"."8层上行呼梯按钮指示灯" )
   END_RUNG
   RUNG wire#powerrail
      N_Contact(operand := #"8层上行呼梯按钮", bit := #连接86)
   END_RUNG wire#w13
   RUNG wire#powerrail
      P_Contact(operand := #"8层下行呼梯按钮", bit := #连接87)
      wire#w14
      S_Coil( "输出"."8层下行呼梯按钮指示灯" )
   END_RUNG
   RUNG wire#powerrail
      N_Contact(operand := #"8层下行呼梯按钮", bit := #连接88)
   END_RUNG wire#w14
   RUNG wire#powerrail
      P_Contact(operand := #"9层上行呼梯按钮", bit := #连接89)
      wire#w15
      S_Coil( "输出"."9层上行呼梯按钮指示灯" )
   END_RUNG
   RUNG wire#powerrail
      N_Contact(operand := #"9层上行呼梯按钮", bit := #连接90)
   END_RUNG wire#w15
   RUNG wire#powerrail
      P_Contact(operand := #"9层下行呼梯按钮", bit := #连接91)
      wire#w16
      S_Coil( "输出"."9层下行呼梯按钮指示灯" )
   END_RUNG
   RUNG wire#powerrail
      N_Contact(operand := #"9层下行呼梯按钮", bit := #连接92)
   END_RUNG wire#w16
   // the same network as SCL:
   #_w1 := #"2层上行呼梯按钮" AND NOT #连接13;   // rising edge of #"2层上行呼梯按钮"
   #连接13 := #"2层上行呼梯按钮";
   #_w2 := NOT #"2层上行呼梯按钮" AND #连接14;   // falling edge of #"2层上行呼梯按钮"
   #连接14 := #"2层上行呼梯按钮";
   IF #_w1 OR #_w2 THEN "输出"."2层上行呼梯按钮指示灯" := TRUE; END_IF;
   #_w3 := #"2层下行呼梯按钮" AND NOT #连接15;   // rising edge of #"2层下行呼梯按钮"
   #连接15 := #"2层下行呼梯按钮";
   #_w4 := NOT #"2层下行呼梯按钮" AND #连接16;   // falling edge of #"2层下行呼梯按钮"
   #连接16 := #"2层下行呼梯按钮";
   IF #_w3 OR #_w4 THEN "输出"."2层下行呼梯按钮指示灯" := TRUE; END_IF;
   #_w5 := #"3层上行呼梯按钮" AND NOT #连接18;   // rising edge of #"3层上行呼梯按钮"
   #连接18 := #"3层上行呼梯按钮";
   #_w6 := NOT #"3层上行呼梯按钮" AND #连接19;   // falling edge of #"3层上行呼梯按钮"
   #连接19 := #"3层上行呼梯按钮";
   IF #_w5 OR #_w6 THEN "输出"."3层上行呼梯按钮指示灯" := TRUE; END_IF;
   #_w7 := #"3层下行呼梯按钮" AND NOT #连接20;   // rising edge of #"3层下行呼梯按钮"
   #连接20 := #"3层下行呼梯按钮";
   #_w8 := NOT #"3层下行呼梯按钮" AND #连接21;   // falling edge of #"3层下行呼梯按钮"
   #连接21 := #"3层下行呼梯按钮";
   IF #_w7 OR #_w8 THEN "输出"."3层下行呼梯按钮指示灯" := TRUE; END_IF;
   #_w9 := #"4层上行呼梯按钮" AND NOT #连接23;   // rising edge of #"4层上行呼梯按钮"
   #连接23 := #"4层上行呼梯按钮";
   #_w10 := NOT #"4层上行呼梯按钮" AND #连接24;   // falling edge of #"4层上行呼梯按钮"
   #连接24 := #"4层上行呼梯按钮";
   IF #_w9 OR #_w10 THEN "输出"."4层上行呼梯按钮指示灯" := TRUE; END_IF;
   #_w11 := #"4层下行呼梯按钮" AND NOT #连接25;   // rising edge of #"4层下行呼梯按钮"
   #连接25 := #"4层下行呼梯按钮";
   #_w12 := NOT #"4层下行呼梯按钮" AND #连接26;   // falling edge of #"4层下行呼梯按钮"
   #连接26 := #"4层下行呼梯按钮";
   IF #_w11 OR #_w12 THEN "输出"."4层下行呼梯按钮指示灯" := TRUE; END_IF;
   #_w13 := #"5层上行呼梯按钮" AND NOT #连接28;   // rising edge of #"5层上行呼梯按钮"
   #连接28 := #"5层上行呼梯按钮";
   #_w14 := NOT #"5层上行呼梯按钮" AND #连接29;   // falling edge of #"5层上行呼梯按钮"
   #连接29 := #"5层上行呼梯按钮";
   IF #_w13 OR #_w14 THEN "输出"."5层上行呼梯按钮指示灯" := TRUE; END_IF;
   #_w15 := #"5层下行呼梯按钮" AND NOT #连接30;   // rising edge of #"5层下行呼梯按钮"
   #连接30 := #"5层下行呼梯按钮";
   #_w16 := NOT #"5层下行呼梯按钮" AND #连接31;   // falling edge of #"5层下行呼梯按钮"
   #连接31 := #"5层下行呼梯按钮";
   IF #_w15 OR #_w16 THEN "输出"."5层下行呼梯按钮指示灯" := TRUE; END_IF;
   #_w17 := #"6层上行呼梯按钮" AND NOT #连接77;   // rising edge of #"6层上行呼梯按钮"
   #连接77 := #"6层上行呼梯按钮";
   #_w18 := NOT #"6层上行呼梯按钮" AND #连接78;   // falling edge of #"6层上行呼梯按钮"
   #连接78 := #"6层上行呼梯按钮";
   IF #_w17 OR #_w18 THEN "输出"."6层上行呼梯按钮指示灯" := TRUE; END_IF;
   #_w19 := #"6层下行呼梯按钮" AND NOT #连接79;   // rising edge of #"6层下行呼梯按钮"
   #连接79 := #"6层下行呼梯按钮";
   #_w20 := NOT #"6层下行呼梯按钮" AND #连接80;   // falling edge of #"6层下行呼梯按钮"
   #连接80 := #"6层下行呼梯按钮";
   IF #_w19 OR #_w20 THEN "输出"."6层下行呼梯按钮指示灯" := TRUE; END_IF;
   #_w21 := #"7层上行呼梯按钮" AND NOT #连接81;   // rising edge of #"7层上行呼梯按钮"
   #连接81 := #"7层上行呼梯按钮";
   #_w22 := NOT #"7层上行呼梯按钮" AND #连接82;   // falling edge of #"7层上行呼梯按钮"
   #连接82 := #"7层上行呼梯按钮";
   IF #_w21 OR #_w22 THEN "输出"."7层上行呼梯按钮指示灯" := TRUE; END_IF;
   #_w23 := #"7层下行呼梯按钮" AND NOT #连接83;   // rising edge of #"7层下行呼梯按钮"
   #连接83 := #"7层下行呼梯按钮";
   #_w24 := NOT #"7层下行呼梯按钮" AND #连接84;   // falling edge of #"7层下行呼梯按钮"
   #连接84 := #"7层下行呼梯按钮";
   IF #_w23 OR #_w24 THEN "输出"."7层下行呼梯按钮指示灯" := TRUE; END_IF;
   #_w25 := #"8层上行呼梯按钮" AND NOT #连接85;   // rising edge of #"8层上行呼梯按钮"
   #连接85 := #"8层上行呼梯按钮";
   #_w26 := NOT #"8层上行呼梯按钮" AND #连接86;   // falling edge of #"8层上行呼梯按钮"
   #连接86 := #"8层上行呼梯按钮";
   IF #_w25 OR #_w26 THEN "输出"."8层上行呼梯按钮指示灯" := TRUE; END_IF;
   #_w27 := #"8层下行呼梯按钮" AND NOT #连接87;   // rising edge of #"8层下行呼梯按钮"
   #连接87 := #"8层下行呼梯按钮";
   #_w28 := NOT #"8层下行呼梯按钮" AND #连接88;   // falling edge of #"8层下行呼梯按钮"
   #连接88 := #"8层下行呼梯按钮";
   IF #_w27 OR #_w28 THEN "输出"."8层下行呼梯按钮指示灯" := TRUE; END_IF;
   #_w29 := #"9层上行呼梯按钮" AND NOT #连接89;   // rising edge of #"9层上行呼梯按钮"
   #连接89 := #"9层上行呼梯按钮";
   #_w30 := NOT #"9层上行呼梯按钮" AND #连接90;   // falling edge of #"9层上行呼梯按钮"
   #连接90 := #"9层上行呼梯按钮";
   IF #_w29 OR #_w30 THEN "输出"."9层上行呼梯按钮指示灯" := TRUE; END_IF;
   #_w31 := #"9层下行呼梯按钮" AND NOT #连接91;   // rising edge of #"9层下行呼梯按钮"
   #连接91 := #"9层下行呼梯按钮";
   #_w32 := NOT #"9层下行呼梯按钮" AND #连接92;   // falling edge of #"9层下行呼梯按钮"
   #连接92 := #"9层下行呼梯按钮";
   IF #_w31 OR #_w32 THEN "输出"."9层下行呼梯按钮指示灯" := TRUE; END_IF;
END_REGION

REGION Network 7: 内呼 按钮与指示灯
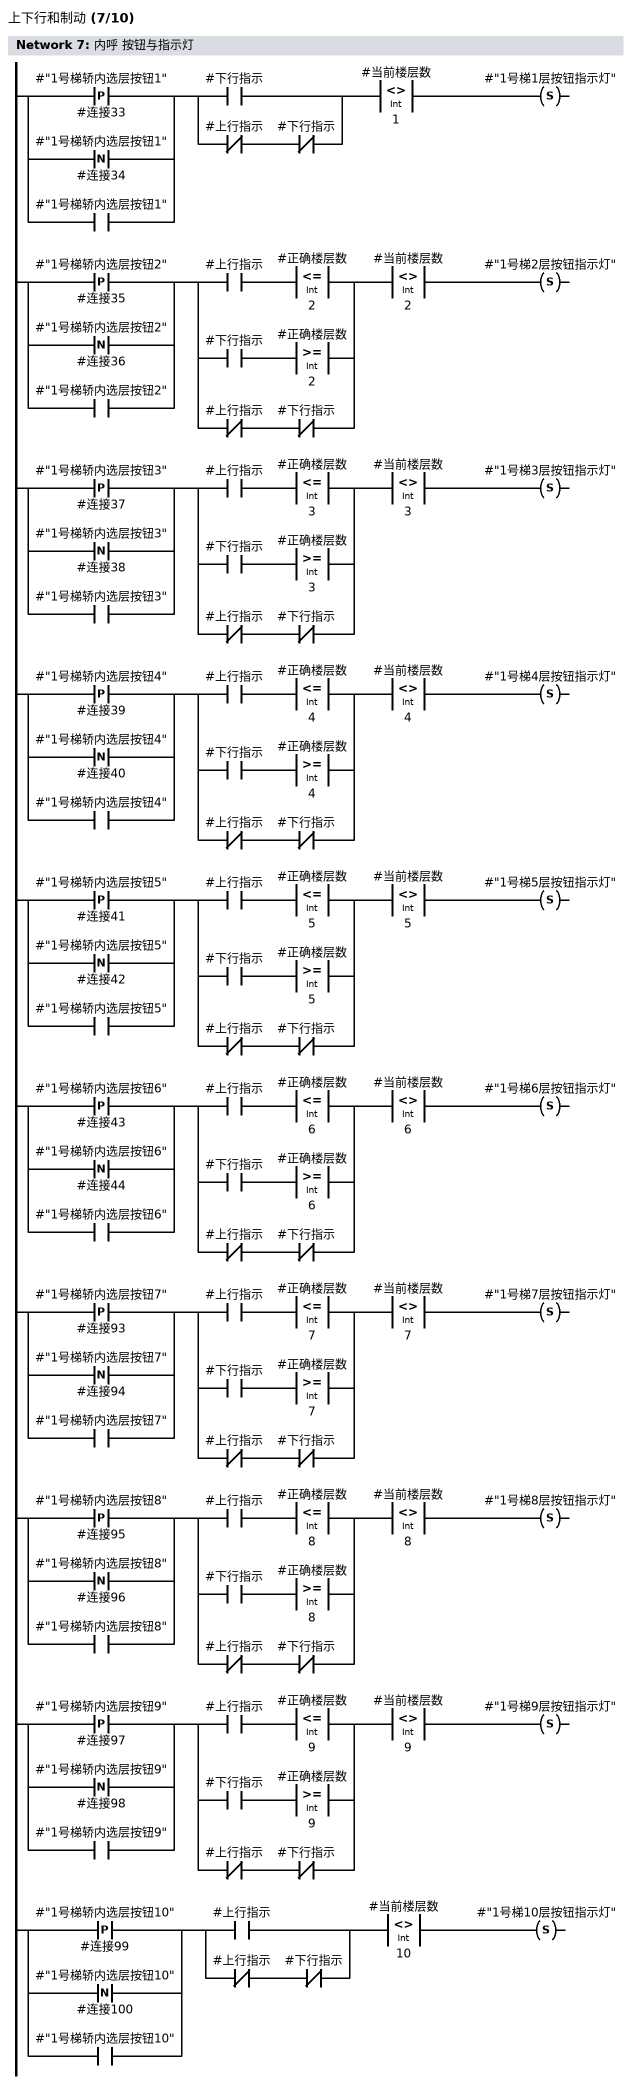
   RUNG wire#powerrail
      P_Contact(operand := #"1号梯轿内选层按钮1", bit := #连接33)
      wire#w1
      Contact( #下行指示 )
      wire#w2
      { S7_Templates := "SrcType := Int" } NE_Contact(in1 := #当前楼层数, in2 := 1)
      S_Coil( #"1号梯1层按钮指示灯" )
   END_RUNG
   RUNG wire#powerrail
      N_Contact(operand := #"1号梯轿内选层按钮1", bit := #连接34)
   END_RUNG wire#w1
   RUNG wire#powerrail
      Contact( #"1号梯轿内选层按钮1" )
   END_RUNG wire#w1
   RUNG wire#w1
      I_Contact( #上行指示 )
      I_Contact( #下行指示 )
   END_RUNG wire#w2
   RUNG wire#powerrail
      P_Contact(operand := #"1号梯轿内选层按钮2", bit := #连接35)
      wire#w3
      Contact( #上行指示 )
      { S7_Templates := "SrcType := Int" } LE_Contact(in1 := #正确楼层数, in2 := 2)
      wire#w4
      { S7_Templates := "SrcType := Int" } NE_Contact(in1 := #当前楼层数, in2 := 2)
      S_Coil( #"1号梯2层按钮指示灯" )
   END_RUNG
   RUNG wire#powerrail
      N_Contact(operand := #"1号梯轿内选层按钮2", bit := #连接36)
   END_RUNG wire#w3
   RUNG wire#powerrail
      Contact( #"1号梯轿内选层按钮2" )
   END_RUNG wire#w3
   RUNG wire#w3
      Contact( #下行指示 )
      { S7_Templates := "SrcType := Int" } GE_Contact(in1 := #正确楼层数, in2 := 2)
   END_RUNG wire#w4
   RUNG wire#w3
      I_Contact( #上行指示 )
      I_Contact( #下行指示 )
   END_RUNG wire#w4
   RUNG wire#powerrail
      P_Contact(operand := #"1号梯轿内选层按钮3", bit := #连接37)
      wire#w5
      Contact( #上行指示 )
      { S7_Templates := "SrcType := Int" } LE_Contact(in1 := #正确楼层数, in2 := 3)
      wire#w6
      { S7_Templates := "SrcType := Int" } NE_Contact(in1 := #当前楼层数, in2 := 3)
      S_Coil( #"1号梯3层按钮指示灯" )
   END_RUNG
   RUNG wire#powerrail
      N_Contact(operand := #"1号梯轿内选层按钮3", bit := #连接38)
   END_RUNG wire#w5
   RUNG wire#powerrail
      Contact( #"1号梯轿内选层按钮3" )
   END_RUNG wire#w5
   RUNG wire#w5
      Contact( #下行指示 )
      { S7_Templates := "SrcType := Int" } GE_Contact(in1 := #正确楼层数, in2 := 3)
   END_RUNG wire#w6
   RUNG wire#w5
      I_Contact( #上行指示 )
      I_Contact( #下行指示 )
   END_RUNG wire#w6
   RUNG wire#powerrail
      P_Contact(operand := #"1号梯轿内选层按钮4", bit := #连接39)
      wire#w7
      Contact( #上行指示 )
      { S7_Templates := "SrcType := Int" } LE_Contact(in1 := #正确楼层数, in2 := 4)
      wire#w8
      { S7_Templates := "SrcType := Int" } NE_Contact(in1 := #当前楼层数, in2 := 4)
      S_Coil( #"1号梯4层按钮指示灯" )
   END_RUNG
   RUNG wire#powerrail
      N_Contact(operand := #"1号梯轿内选层按钮4", bit := #连接40)
   END_RUNG wire#w7
   RUNG wire#powerrail
      Contact( #"1号梯轿内选层按钮4" )
   END_RUNG wire#w7
   RUNG wire#w7
      Contact( #下行指示 )
      { S7_Templates := "SrcType := Int" } GE_Contact(in1 := #正确楼层数, in2 := 4)
   END_RUNG wire#w8
   RUNG wire#w7
      I_Contact( #上行指示 )
      I_Contact( #下行指示 )
   END_RUNG wire#w8
   RUNG wire#powerrail
      P_Contact(operand := #"1号梯轿内选层按钮5", bit := #连接41)
      wire#w9
      Contact( #上行指示 )
      { S7_Templates := "SrcType := Int" } LE_Contact(in1 := #正确楼层数, in2 := 5)
      wire#w10
      { S7_Templates := "SrcType := Int" } NE_Contact(in1 := #当前楼层数, in2 := 5)
      S_Coil( #"1号梯5层按钮指示灯" )
   END_RUNG
   RUNG wire#powerrail
      N_Contact(operand := #"1号梯轿内选层按钮5", bit := #连接42)
   END_RUNG wire#w9
   RUNG wire#powerrail
      Contact( #"1号梯轿内选层按钮5" )
   END_RUNG wire#w9
   RUNG wire#w9
      Contact( #下行指示 )
      { S7_Templates := "SrcType := Int" } GE_Contact(in1 := #正确楼层数, in2 := 5)
   END_RUNG wire#w10
   RUNG wire#w9
      I_Contact( #上行指示 )
      I_Contact( #下行指示 )
   END_RUNG wire#w10
   RUNG wire#powerrail
      P_Contact(operand := #"1号梯轿内选层按钮6", bit := #连接43)
      wire#w11
      Contact( #上行指示 )
      { S7_Templates := "SrcType := Int" } LE_Contact(in1 := #正确楼层数, in2 := 6)
      wire#w12
      { S7_Templates := "SrcType := Int" } NE_Contact(in1 := #当前楼层数, in2 := 6)
      S_Coil( #"1号梯6层按钮指示灯" )
   END_RUNG
   RUNG wire#powerrail
      N_Contact(operand := #"1号梯轿内选层按钮6", bit := #连接44)
   END_RUNG wire#w11
   RUNG wire#powerrail
      Contact( #"1号梯轿内选层按钮6" )
   END_RUNG wire#w11
   RUNG wire#w11
      Contact( #下行指示 )
      { S7_Templates := "SrcType := Int" } GE_Contact(in1 := #正确楼层数, in2 := 6)
   END_RUNG wire#w12
   RUNG wire#w11
      I_Contact( #上行指示 )
      I_Contact( #下行指示 )
   END_RUNG wire#w12
   RUNG wire#powerrail
      P_Contact(operand := #"1号梯轿内选层按钮7", bit := #连接93)
      wire#w13
      Contact( #上行指示 )
      { S7_Templates := "SrcType := Int" } LE_Contact(in1 := #正确楼层数, in2 := 7)
      wire#w14
      { S7_Templates := "SrcType := Int" } NE_Contact(in1 := #当前楼层数, in2 := 7)
      S_Coil( #"1号梯7层按钮指示灯" )
   END_RUNG
   RUNG wire#powerrail
      N_Contact(operand := #"1号梯轿内选层按钮7", bit := #连接94)
   END_RUNG wire#w13
   RUNG wire#powerrail
      Contact( #"1号梯轿内选层按钮7" )
   END_RUNG wire#w13
   RUNG wire#w13
      Contact( #下行指示 )
      { S7_Templates := "SrcType := Int" } GE_Contact(in1 := #正确楼层数, in2 := 7)
   END_RUNG wire#w14
   RUNG wire#w13
      I_Contact( #上行指示 )
      I_Contact( #下行指示 )
   END_RUNG wire#w14
   RUNG wire#powerrail
      P_Contact(operand := #"1号梯轿内选层按钮8", bit := #连接95)
      wire#w15
      Contact( #上行指示 )
      { S7_Templates := "SrcType := Int" } LE_Contact(in1 := #正确楼层数, in2 := 8)
      wire#w16
      { S7_Templates := "SrcType := Int" } NE_Contact(in1 := #当前楼层数, in2 := 8)
      S_Coil( #"1号梯8层按钮指示灯" )
   END_RUNG
   RUNG wire#powerrail
      N_Contact(operand := #"1号梯轿内选层按钮8", bit := #连接96)
   END_RUNG wire#w15
   RUNG wire#powerrail
      Contact( #"1号梯轿内选层按钮8" )
   END_RUNG wire#w15
   RUNG wire#w15
      Contact( #下行指示 )
      { S7_Templates := "SrcType := Int" } GE_Contact(in1 := #正确楼层数, in2 := 8)
   END_RUNG wire#w16
   RUNG wire#w15
      I_Contact( #上行指示 )
      I_Contact( #下行指示 )
   END_RUNG wire#w16
   RUNG wire#powerrail
      P_Contact(operand := #"1号梯轿内选层按钮9", bit := #连接97)
      wire#w17
      Contact( #上行指示 )
      { S7_Templates := "SrcType := Int" } LE_Contact(in1 := #正确楼层数, in2 := 9)
      wire#w18
      { S7_Templates := "SrcType := Int" } NE_Contact(in1 := #当前楼层数, in2 := 9)
      S_Coil( #"1号梯9层按钮指示灯" )
   END_RUNG
   RUNG wire#powerrail
      N_Contact(operand := #"1号梯轿内选层按钮9", bit := #连接98)
   END_RUNG wire#w17
   RUNG wire#powerrail
      Contact( #"1号梯轿内选层按钮9" )
   END_RUNG wire#w17
   RUNG wire#w17
      Contact( #下行指示 )
      { S7_Templates := "SrcType := Int" } GE_Contact(in1 := #正确楼层数, in2 := 9)
   END_RUNG wire#w18
   RUNG wire#w17
      I_Contact( #上行指示 )
      I_Contact( #下行指示 )
   END_RUNG wire#w18
   RUNG wire#powerrail
      P_Contact(operand := #"1号梯轿内选层按钮10", bit := #连接99)
      wire#w19
      Contact( #上行指示 )
      wire#w20
      { S7_Templates := "SrcType := Int" } NE_Contact(in1 := #当前楼层数, in2 := 10)
      S_Coil( #"1号梯10层按钮指示灯" )
   END_RUNG
   RUNG wire#powerrail
      N_Contact(operand := #"1号梯轿内选层按钮10", bit := #连接100)
   END_RUNG wire#w19
   RUNG wire#powerrail
      Contact( #"1号梯轿内选层按钮10" )
   END_RUNG wire#w19
   RUNG wire#w19
      I_Contact( #上行指示 )
      I_Contact( #下行指示 )
   END_RUNG wire#w20
   // the same network as SCL:
   #_w1 := #"1号梯轿内选层按钮1" AND NOT #连接33;   // rising edge of #"1号梯轿内选层按钮1"
   #连接33 := #"1号梯轿内选层按钮1";
   #_w2 := NOT #"1号梯轿内选层按钮1" AND #连接34;   // falling edge of #"1号梯轿内选层按钮1"
   #连接34 := #"1号梯轿内选层按钮1";
   IF (#_w1 OR #_w2 OR #"1号梯轿内选层按钮1") AND (#下行指示 OR (NOT #上行指示 AND NOT #下行指示)) AND (#当前楼层数 <> 1) THEN
       #"1号梯1层按钮指示灯" := TRUE;
   END_IF;
   #_w3 := #"1号梯轿内选层按钮2" AND NOT #连接35;   // rising edge of #"1号梯轿内选层按钮2"
   #连接35 := #"1号梯轿内选层按钮2";
   #_w4 := NOT #"1号梯轿内选层按钮2" AND #连接36;   // falling edge of #"1号梯轿内选层按钮2"
   #连接36 := #"1号梯轿内选层按钮2";
   IF (#_w3 OR #_w4 OR #"1号梯轿内选层按钮2") AND ((#上行指示 AND (#正确楼层数 <= 2)) OR (#下行指示 AND (#正确楼层数 >= 2)) OR (NOT #上行指示 AND NOT #下行指示)) AND (#当前楼层数 <> 2) THEN
       #"1号梯2层按钮指示灯" := TRUE;
   END_IF;
   #_w5 := #"1号梯轿内选层按钮3" AND NOT #连接37;   // rising edge of #"1号梯轿内选层按钮3"
   #连接37 := #"1号梯轿内选层按钮3";
   #_w6 := NOT #"1号梯轿内选层按钮3" AND #连接38;   // falling edge of #"1号梯轿内选层按钮3"
   #连接38 := #"1号梯轿内选层按钮3";
   IF (#_w5 OR #_w6 OR #"1号梯轿内选层按钮3") AND ((#上行指示 AND (#正确楼层数 <= 3)) OR (#下行指示 AND (#正确楼层数 >= 3)) OR (NOT #上行指示 AND NOT #下行指示)) AND (#当前楼层数 <> 3) THEN
       #"1号梯3层按钮指示灯" := TRUE;
   END_IF;
   #_w7 := #"1号梯轿内选层按钮4" AND NOT #连接39;   // rising edge of #"1号梯轿内选层按钮4"
   #连接39 := #"1号梯轿内选层按钮4";
   #_w8 := NOT #"1号梯轿内选层按钮4" AND #连接40;   // falling edge of #"1号梯轿内选层按钮4"
   #连接40 := #"1号梯轿内选层按钮4";
   IF (#_w7 OR #_w8 OR #"1号梯轿内选层按钮4") AND ((#上行指示 AND (#正确楼层数 <= 4)) OR (#下行指示 AND (#正确楼层数 >= 4)) OR (NOT #上行指示 AND NOT #下行指示)) AND (#当前楼层数 <> 4) THEN
       #"1号梯4层按钮指示灯" := TRUE;
   END_IF;
   #_w9 := #"1号梯轿内选层按钮5" AND NOT #连接41;   // rising edge of #"1号梯轿内选层按钮5"
   #连接41 := #"1号梯轿内选层按钮5";
   #_w10 := NOT #"1号梯轿内选层按钮5" AND #连接42;   // falling edge of #"1号梯轿内选层按钮5"
   #连接42 := #"1号梯轿内选层按钮5";
   IF (#_w9 OR #_w10 OR #"1号梯轿内选层按钮5") AND ((#上行指示 AND (#正确楼层数 <= 5)) OR (#下行指示 AND (#正确楼层数 >= 5)) OR (NOT #上行指示 AND NOT #下行指示)) AND (#当前楼层数 <> 5) THEN
       #"1号梯5层按钮指示灯" := TRUE;
   END_IF;
   #_w11 := #"1号梯轿内选层按钮6" AND NOT #连接43;   // rising edge of #"1号梯轿内选层按钮6"
   #连接43 := #"1号梯轿内选层按钮6";
   #_w12 := NOT #"1号梯轿内选层按钮6" AND #连接44;   // falling edge of #"1号梯轿内选层按钮6"
   #连接44 := #"1号梯轿内选层按钮6";
   IF (#_w11 OR #_w12 OR #"1号梯轿内选层按钮6") AND ((#上行指示 AND (#正确楼层数 <= 6)) OR (#下行指示 AND (#正确楼层数 >= 6)) OR (NOT #上行指示 AND NOT #下行指示)) AND (#当前楼层数 <> 6) THEN
       #"1号梯6层按钮指示灯" := TRUE;
   END_IF;
   #_w13 := #"1号梯轿内选层按钮7" AND NOT #连接93;   // rising edge of #"1号梯轿内选层按钮7"
   #连接93 := #"1号梯轿内选层按钮7";
   #_w14 := NOT #"1号梯轿内选层按钮7" AND #连接94;   // falling edge of #"1号梯轿内选层按钮7"
   #连接94 := #"1号梯轿内选层按钮7";
   IF (#_w13 OR #_w14 OR #"1号梯轿内选层按钮7") AND ((#上行指示 AND (#正确楼层数 <= 7)) OR (#下行指示 AND (#正确楼层数 >= 7)) OR (NOT #上行指示 AND NOT #下行指示)) AND (#当前楼层数 <> 7) THEN
       #"1号梯7层按钮指示灯" := TRUE;
   END_IF;
   #_w15 := #"1号梯轿内选层按钮8" AND NOT #连接95;   // rising edge of #"1号梯轿内选层按钮8"
   #连接95 := #"1号梯轿内选层按钮8";
   #_w16 := NOT #"1号梯轿内选层按钮8" AND #连接96;   // falling edge of #"1号梯轿内选层按钮8"
   #连接96 := #"1号梯轿内选层按钮8";
   IF (#_w15 OR #_w16 OR #"1号梯轿内选层按钮8") AND ((#上行指示 AND (#正确楼层数 <= 8)) OR (#下行指示 AND (#正确楼层数 >= 8)) OR (NOT #上行指示 AND NOT #下行指示)) AND (#当前楼层数 <> 8) THEN
       #"1号梯8层按钮指示灯" := TRUE;
   END_IF;
   #_w17 := #"1号梯轿内选层按钮9" AND NOT #连接97;   // rising edge of #"1号梯轿内选层按钮9"
   #连接97 := #"1号梯轿内选层按钮9";
   #_w18 := NOT #"1号梯轿内选层按钮9" AND #连接98;   // falling edge of #"1号梯轿内选层按钮9"
   #连接98 := #"1号梯轿内选层按钮9";
   IF (#_w17 OR #_w18 OR #"1号梯轿内选层按钮9") AND ((#上行指示 AND (#正确楼层数 <= 9)) OR (#下行指示 AND (#正确楼层数 >= 9)) OR (NOT #上行指示 AND NOT #下行指示)) AND (#当前楼层数 <> 9) THEN
       #"1号梯9层按钮指示灯" := TRUE;
   END_IF;
   #_w19 := #"1号梯轿内选层按钮10" AND NOT #连接99;   // rising edge of #"1号梯轿内选层按钮10"
   #连接99 := #"1号梯轿内选层按钮10";
   #_w20 := NOT #"1号梯轿内选层按钮10" AND #连接100;   // falling edge of #"1号梯轿内选层按钮10"
   #连接100 := #"1号梯轿内选层按钮10";
   IF (#_w19 OR #_w20 OR #"1号梯轿内选层按钮10") AND (#上行指示 OR (NOT #上行指示 AND NOT #下行指示)) AND (#当前楼层数 <> 10) THEN
       #"1号梯10层按钮指示灯" := TRUE;
   END_IF;
END_REGION

REGION Network 8: 灭灯 （按上下行顺序）
   // 到达1，10层后内置按钮清零
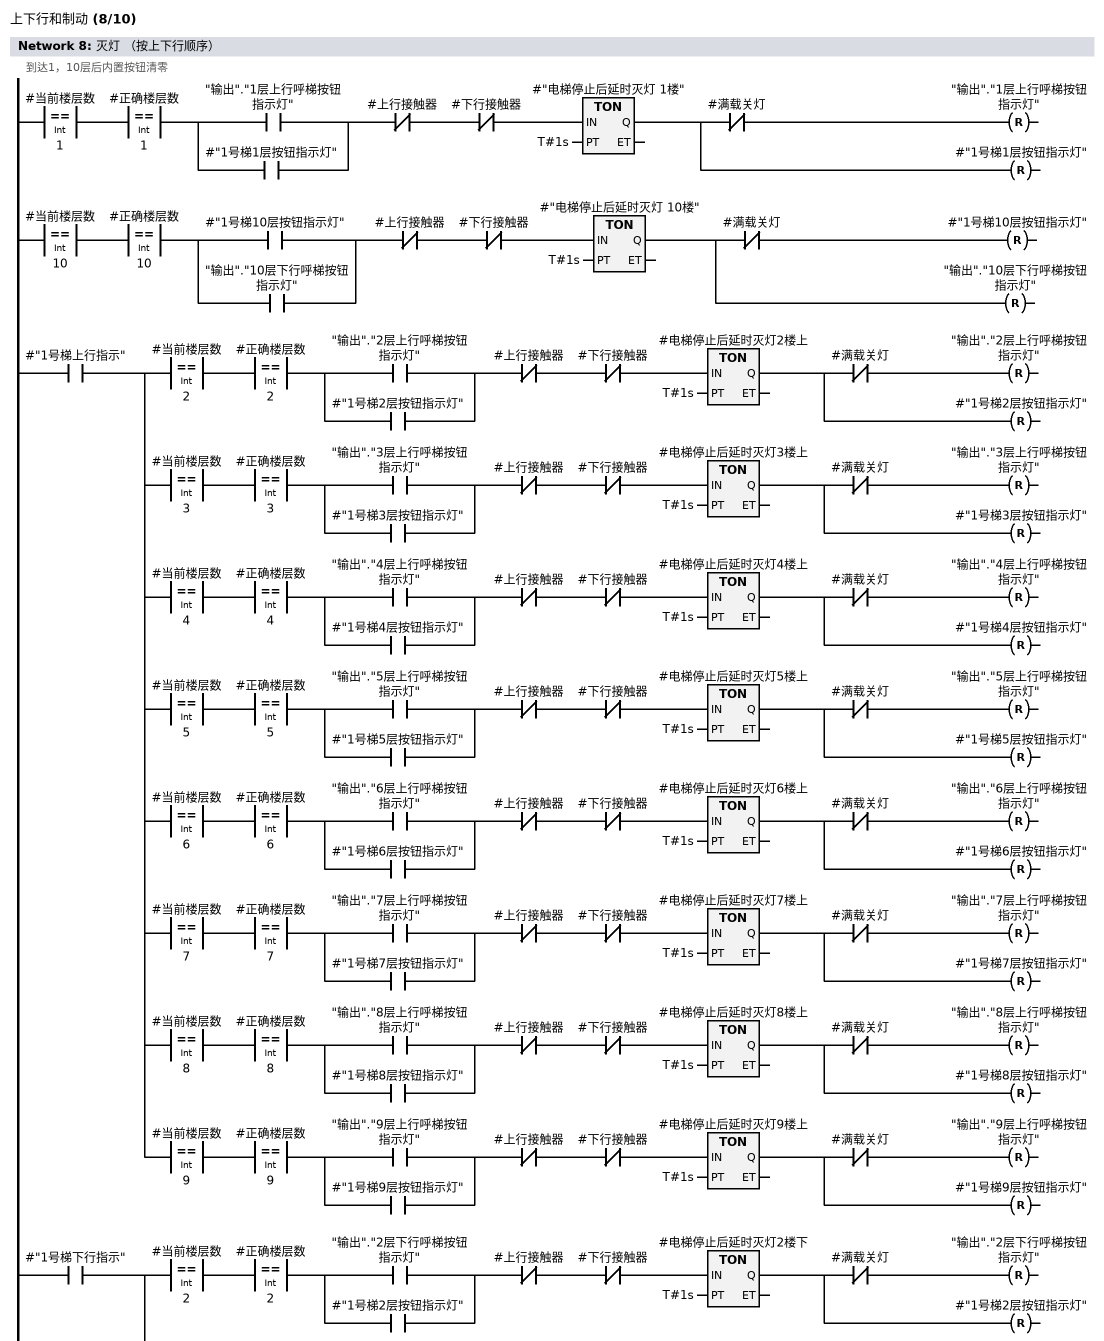
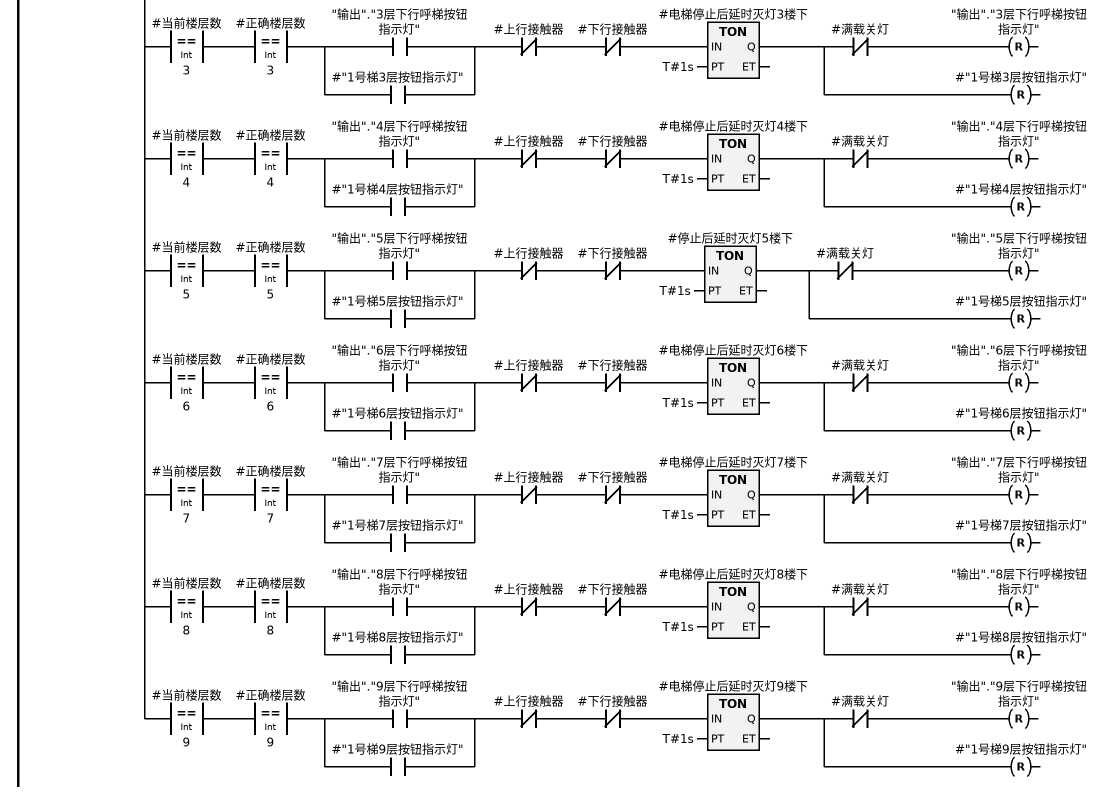
   #"电梯停止后延时灭灯 1楼"(IN := (#当前楼层数 = 1) AND (#正确楼层数 = 1) AND ("输出"."1层上行呼梯按钮指示灯" OR #"1号梯1层按钮指示灯") AND NOT #上行接触器 AND NOT #下行接触器,   // TON
                   PT := T#1s);
   IF #"电梯停止后延时灭灯 1楼".Q AND NOT #满载关灯 THEN "输出"."1层上行呼梯按钮指示灯" := FALSE; END_IF;
   IF #"电梯停止后延时灭灯 1楼".Q THEN #"1号梯1层按钮指示灯" := FALSE; END_IF;
   #"电梯停止后延时灭灯 10楼"(IN := (#当前楼层数 = 10) AND (#正确楼层数 = 10) AND (#"1号梯10层按钮指示灯" OR "输出"."10层下行呼梯按钮指示灯") AND NOT #上行接触器 AND NOT #下行接触器,   // TON
                    PT := T#1s);
   IF #"电梯停止后延时灭灯 10楼".Q AND NOT #满载关灯 THEN #"1号梯10层按钮指示灯" := FALSE; END_IF;
   IF #"电梯停止后延时灭灯 10楼".Q THEN "输出"."10层下行呼梯按钮指示灯" := FALSE; END_IF;
   #电梯停止后延时灭灯2楼上(IN := #"1号梯上行指示" AND (#当前楼层数 = 2) AND (#正确楼层数 = 2) AND ("输出"."2层上行呼梯按钮指示灯" OR #"1号梯2层按钮指示灯") AND NOT #上行接触器 AND NOT #下行接触器,   // TON
                 PT := T#1s);
   IF #电梯停止后延时灭灯2楼上.Q AND NOT #满载关灯 THEN "输出"."2层上行呼梯按钮指示灯" := FALSE; END_IF;
   IF #电梯停止后延时灭灯2楼上.Q THEN #"1号梯2层按钮指示灯" := FALSE; END_IF;
   #电梯停止后延时灭灯3楼上(IN := #"1号梯上行指示" AND (#当前楼层数 = 3) AND (#正确楼层数 = 3) AND ("输出"."3层上行呼梯按钮指示灯" OR #"1号梯3层按钮指示灯") AND NOT #上行接触器 AND NOT #下行接触器,   // TON
                 PT := T#1s);
   IF #电梯停止后延时灭灯3楼上.Q AND NOT #满载关灯 THEN "输出"."3层上行呼梯按钮指示灯" := FALSE; END_IF;
   IF #电梯停止后延时灭灯3楼上.Q THEN #"1号梯3层按钮指示灯" := FALSE; END_IF;
   #电梯停止后延时灭灯4楼上(IN := #"1号梯上行指示" AND (#当前楼层数 = 4) AND (#正确楼层数 = 4) AND ("输出"."4层上行呼梯按钮指示灯" OR #"1号梯4层按钮指示灯") AND NOT #上行接触器 AND NOT #下行接触器,   // TON
                 PT := T#1s);
   IF #电梯停止后延时灭灯4楼上.Q AND NOT #满载关灯 THEN "输出"."4层上行呼梯按钮指示灯" := FALSE; END_IF;
   IF #电梯停止后延时灭灯4楼上.Q THEN #"1号梯4层按钮指示灯" := FALSE; END_IF;
   #电梯停止后延时灭灯5楼上(IN := #"1号梯上行指示" AND (#当前楼层数 = 5) AND (#正确楼层数 = 5) AND ("输出"."5层上行呼梯按钮指示灯" OR #"1号梯5层按钮指示灯") AND NOT #上行接触器 AND NOT #下行接触器,   // TON
                 PT := T#1s);
   IF #电梯停止后延时灭灯5楼上.Q AND NOT #满载关灯 THEN "输出"."5层上行呼梯按钮指示灯" := FALSE; END_IF;
   IF #电梯停止后延时灭灯5楼上.Q THEN #"1号梯5层按钮指示灯" := FALSE; END_IF;
   #电梯停止后延时灭灯6楼上(IN := #"1号梯上行指示" AND (#当前楼层数 = 6) AND (#正确楼层数 = 6) AND ("输出"."6层上行呼梯按钮指示灯" OR #"1号梯6层按钮指示灯") AND NOT #上行接触器 AND NOT #下行接触器,   // TON
                 PT := T#1s);
   IF #电梯停止后延时灭灯6楼上.Q AND NOT #满载关灯 THEN "输出"."6层上行呼梯按钮指示灯" := FALSE; END_IF;
   IF #电梯停止后延时灭灯6楼上.Q THEN #"1号梯6层按钮指示灯" := FALSE; END_IF;
   #电梯停止后延时灭灯7楼上(IN := #"1号梯上行指示" AND (#当前楼层数 = 7) AND (#正确楼层数 = 7) AND ("输出"."7层上行呼梯按钮指示灯" OR #"1号梯7层按钮指示灯") AND NOT #上行接触器 AND NOT #下行接触器,   // TON
                 PT := T#1s);
   IF #电梯停止后延时灭灯7楼上.Q AND NOT #满载关灯 THEN "输出"."7层上行呼梯按钮指示灯" := FALSE; END_IF;
   IF #电梯停止后延时灭灯7楼上.Q THEN #"1号梯7层按钮指示灯" := FALSE; END_IF;
   #电梯停止后延时灭灯8楼上(IN := #"1号梯上行指示" AND (#当前楼层数 = 8) AND (#正确楼层数 = 8) AND ("输出"."8层上行呼梯按钮指示灯" OR #"1号梯8层按钮指示灯") AND NOT #上行接触器 AND NOT #下行接触器,   // TON
                 PT := T#1s);
   IF #电梯停止后延时灭灯8楼上.Q AND NOT #满载关灯 THEN "输出"."8层上行呼梯按钮指示灯" := FALSE; END_IF;
   IF #电梯停止后延时灭灯8楼上.Q THEN #"1号梯8层按钮指示灯" := FALSE; END_IF;
   #电梯停止后延时灭灯9楼上(IN := #"1号梯上行指示" AND (#当前楼层数 = 9) AND (#正确楼层数 = 9) AND ("输出"."9层上行呼梯按钮指示灯" OR #"1号梯9层按钮指示灯") AND NOT #上行接触器 AND NOT #下行接触器,   // TON
                 PT := T#1s);
   IF #电梯停止后延时灭灯9楼上.Q AND NOT #满载关灯 THEN "输出"."9层上行呼梯按钮指示灯" := FALSE; END_IF;
   IF #电梯停止后延时灭灯9楼上.Q THEN #"1号梯9层按钮指示灯" := FALSE; END_IF;
   #电梯停止后延时灭灯2楼下(IN := #"1号梯下行指示" AND (#当前楼层数 = 2) AND (#正确楼层数 = 2) AND ("输出"."2层下行呼梯按钮指示灯" OR #"1号梯2层按钮指示灯") AND NOT #上行接触器 AND NOT #下行接触器,   // TON
                 PT := T#1s);
   IF #电梯停止后延时灭灯2楼下.Q AND NOT #满载关灯 THEN "输出"."2层下行呼梯按钮指示灯" := FALSE; END_IF;
   IF #电梯停止后延时灭灯2楼下.Q THEN #"1号梯2层按钮指示灯" := FALSE; END_IF;
   #电梯停止后延时灭灯3楼下(IN := #"1号梯下行指示" AND (#当前楼层数 = 3) AND (#正确楼层数 = 3) AND ("输出"."3层下行呼梯按钮指示灯" OR #"1号梯3层按钮指示灯") AND NOT #上行接触器 AND NOT #下行接触器,   // TON
                 PT := T#1s);
   IF #电梯停止后延时灭灯3楼下.Q AND NOT #满载关灯 THEN "输出"."3层下行呼梯按钮指示灯" := FALSE; END_IF;
   IF #电梯停止后延时灭灯3楼下.Q THEN #"1号梯3层按钮指示灯" := FALSE; END_IF;
   #电梯停止后延时灭灯4楼下(IN := #"1号梯下行指示" AND (#当前楼层数 = 4) AND (#正确楼层数 = 4) AND ("输出"."4层下行呼梯按钮指示灯" OR #"1号梯4层按钮指示灯") AND NOT #上行接触器 AND NOT #下行接触器,   // TON
                 PT := T#1s);
   IF #电梯停止后延时灭灯4楼下.Q AND NOT #满载关灯 THEN "输出"."4层下行呼梯按钮指示灯" := FALSE; END_IF;
   IF #电梯停止后延时灭灯4楼下.Q THEN #"1号梯4层按钮指示灯" := FALSE; END_IF;
   #停止后延时灭灯5楼下(IN := #"1号梯下行指示" AND (#当前楼层数 = 5) AND (#正确楼层数 = 5) AND ("输出"."5层下行呼梯按钮指示灯" OR #"1号梯5层按钮指示灯") AND NOT #上行接触器 AND NOT #下行接触器,   // TON
               PT := T#1s);
   IF #停止后延时灭灯5楼下.Q AND NOT #满载关灯 THEN "输出"."5层下行呼梯按钮指示灯" := FALSE; END_IF;
   IF #停止后延时灭灯5楼下.Q THEN #"1号梯5层按钮指示灯" := FALSE; END_IF;
   #电梯停止后延时灭灯6楼下(IN := #"1号梯下行指示" AND (#当前楼层数 = 6) AND (#正确楼层数 = 6) AND ("输出"."6层下行呼梯按钮指示灯" OR #"1号梯6层按钮指示灯") AND NOT #上行接触器 AND NOT #下行接触器,   // TON
                 PT := T#1s);
   IF #电梯停止后延时灭灯6楼下.Q AND NOT #满载关灯 THEN "输出"."6层下行呼梯按钮指示灯" := FALSE; END_IF;
   IF #电梯停止后延时灭灯6楼下.Q THEN #"1号梯6层按钮指示灯" := FALSE; END_IF;
   #电梯停止后延时灭灯7楼下(IN := #"1号梯下行指示" AND (#当前楼层数 = 7) AND (#正确楼层数 = 7) AND ("输出"."7层下行呼梯按钮指示灯" OR #"1号梯7层按钮指示灯") AND NOT #上行接触器 AND NOT #下行接触器,   // TON
                 PT := T#1s);
   IF #电梯停止后延时灭灯7楼下.Q AND NOT #满载关灯 THEN "输出"."7层下行呼梯按钮指示灯" := FALSE; END_IF;
   IF #电梯停止后延时灭灯7楼下.Q THEN #"1号梯7层按钮指示灯" := FALSE; END_IF;
   #电梯停止后延时灭灯8楼下(IN := #"1号梯下行指示" AND (#当前楼层数 = 8) AND (#正确楼层数 = 8) AND ("输出"."8层下行呼梯按钮指示灯" OR #"1号梯8层按钮指示灯") AND NOT #上行接触器 AND NOT #下行接触器,   // TON
                 PT := T#1s);
   IF #电梯停止后延时灭灯8楼下.Q AND NOT #满载关灯 THEN "输出"."8层下行呼梯按钮指示灯" := FALSE; END_IF;
   IF #电梯停止后延时灭灯8楼下.Q THEN #"1号梯8层按钮指示灯" := FALSE; END_IF;
   #电梯停止后延时灭灯9楼下(IN := #"1号梯下行指示" AND (#当前楼层数 = 9) AND (#正确楼层数 = 9) AND ("输出"."9层下行呼梯按钮指示灯" OR #"1号梯9层按钮指示灯") AND NOT #上行接触器 AND NOT #下行接触器,   // TON
                 PT := T#1s);
   IF #电梯停止后延时灭灯9楼下.Q AND NOT #满载关灯 THEN "输出"."9层下行呼梯按钮指示灯" := FALSE; END_IF;
   IF #电梯停止后延时灭灯9楼下.Q THEN #"1号梯9层按钮指示灯" := FALSE; END_IF;
END_REGION

REGION Network 9: 制动
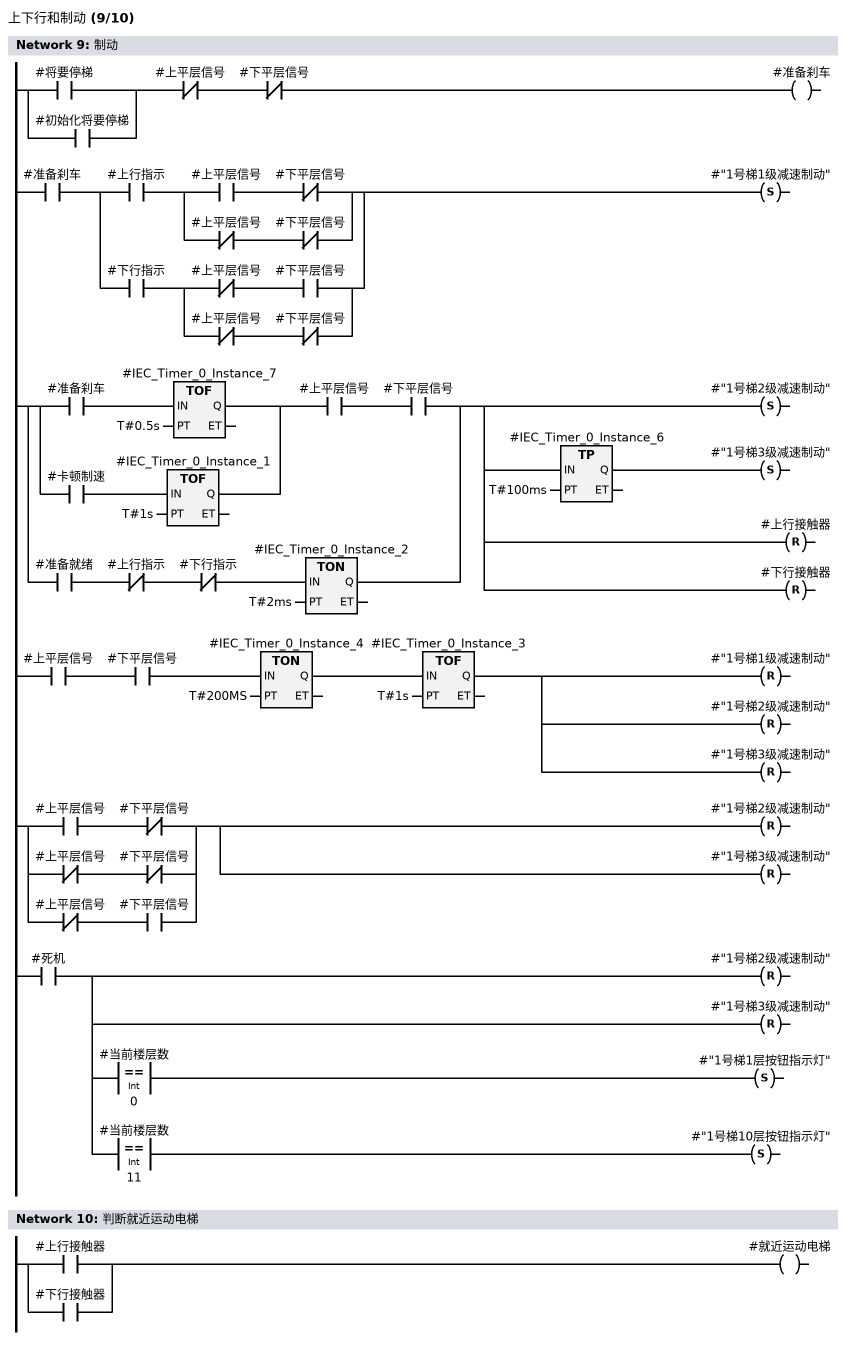
   #准备刹车 := (#将要停梯 OR #初始化将要停梯) AND NOT #上平层信号 AND NOT #下平层信号;
   IF #准备刹车 AND ((#上行指示 AND ((#上平层信号 AND NOT #下平层信号) OR (NOT #上平层信号 AND NOT #下平层信号))) OR (#下行指示 AND ((NOT #上平层信号 AND #下平层信号) OR (NOT #上平层信号 AND NOT #下平层信号)))) THEN
       #"1号梯1级减速制动" := TRUE;
   END_IF;
   #IEC_Timer_0_Instance_7(IN := #准备刹车, PT := T#0.5s);   // TOF
   #IEC_Timer_0_Instance_1(IN := #卡顿制速, PT := T#1s);   // TOF
   #IEC_Timer_0_Instance_2(IN := #准备就绪 AND NOT #上行指示 AND NOT #下行指示, PT := T#2ms);   // TON
   #_w1 := ((#IEC_Timer_0_Instance_7.Q OR #IEC_Timer_0_Instance_1.Q) AND #上平层信号 AND #下平层信号) OR #IEC_Timer_0_Instance_2.Q;
   IF #_w1 THEN #"1号梯2级减速制动" := TRUE; END_IF;
   #IEC_Timer_0_Instance_6(IN := #_w1, PT := T#100ms);   // TP
   IF #IEC_Timer_0_Instance_6.Q THEN #"1号梯3级减速制动" := TRUE; END_IF;
   IF #_w1 THEN
       #上行接触器 := FALSE;
       #下行接触器 := FALSE;
   END_IF;
   #IEC_Timer_0_Instance_4(IN := #上平层信号 AND #下平层信号, PT := T#200MS);   // TON
   #IEC_Timer_0_Instance_3(IN := #IEC_Timer_0_Instance_4.Q, PT := T#1s);   // TOF
   IF #IEC_Timer_0_Instance_3.Q THEN
       #"1号梯1级减速制动" := FALSE;
       #"1号梯2级减速制动" := FALSE;
       #"1号梯3级减速制动" := FALSE;
   END_IF;
   IF (#上平层信号 AND NOT #下平层信号) OR (NOT #上平层信号 AND NOT #下平层信号) OR (NOT #上平层信号 AND #下平层信号) THEN
       #"1号梯2级减速制动" := FALSE;
       #"1号梯3级减速制动" := FALSE;
   END_IF;
   IF #死机 THEN
       #"1号梯2级减速制动" := FALSE;
       #"1号梯3级减速制动" := FALSE;
   END_IF;
   IF #死机 AND (#当前楼层数 = 0) THEN #"1号梯1层按钮指示灯" := TRUE; END_IF;
   IF #死机 AND (#当前楼层数 = 11) THEN #"1号梯10层按钮指示灯" := TRUE; END_IF;
END_REGION

REGION Network 10: 判断就近运动电梯
   RUNG wire#powerrail
      Contact( #上行接触器 )
      wire#w1
      Coil( #就近运动电梯 )
   END_RUNG
   RUNG wire#powerrail
      Contact( #下行接触器 )
   END_RUNG wire#w1
   // the same network as SCL:
   #就近运动电梯 := #上行接触器 OR #下行接触器;
END_REGION

REGION Network 11: 判断是否满载
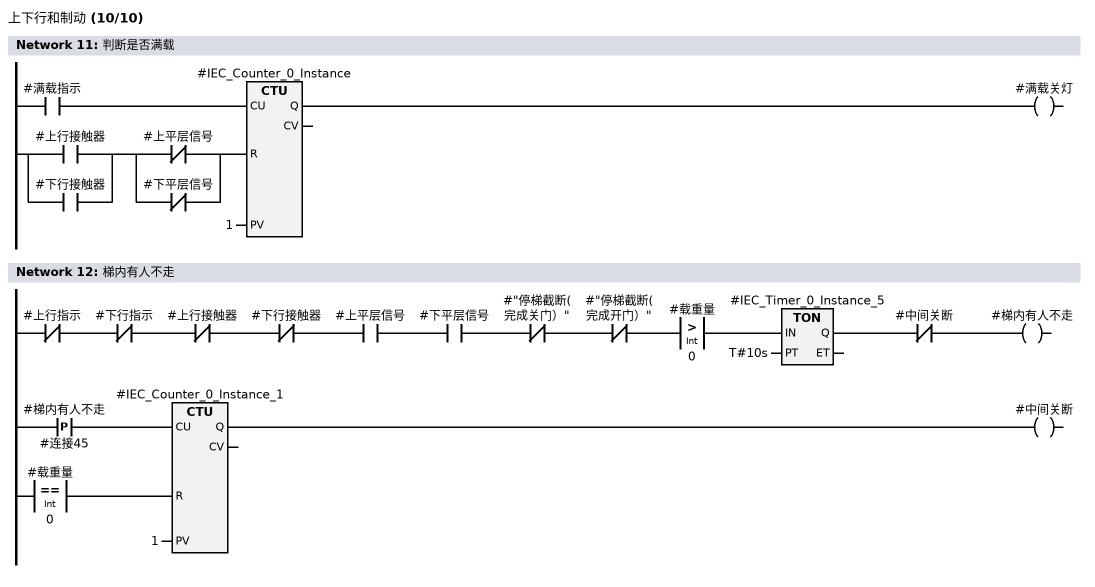
   #IEC_Counter_0_Instance(CU := #满载指示, R := (#上行接触器 OR #下行接触器) AND (NOT #上平层信号 OR NOT #下平层信号), PV := 1);   // CTU
   #满载关灯 := #IEC_Counter_0_Instance.Q;
END_REGION

REGION Network 12: 梯内有人不走
   #IEC_Timer_0_Instance_5(IN := NOT #上行指示 AND NOT #下行指示 AND NOT #上行接触器 AND NOT #下行接触器 AND #上平层信号 AND #下平层信号 AND NOT #"停梯截断(完成关门）" AND NOT #"停梯截断(完成开门）" AND (#载重量 > 0),   // TON
                           PT := T#10s);
   #梯内有人不走 := #IEC_Timer_0_Instance_5.Q AND NOT #中间关断;
   #_w1 := #梯内有人不走 AND NOT #连接45;   // rising edge of #梯内有人不走
   #连接45 := #梯内有人不走;
   #IEC_Counter_0_Instance_1(CU := #_w1, R := #载重量 = 0, PV := 1);   // CTU
   #中间关断 := #IEC_Counter_0_Instance_1.Q;
END_REGION
END_FUNCTION_BLOCK

FUNCTION_BLOCK "优先级响应开关门"   // FB11, LAD
{ S7_Optimized_Access := 'TRUE' }
VERSION : 0.1
   VAR_INPUT
      准备就绪 : Bool;
      "1号梯转换后载重量" : Int;
      "1号梯上行指示" : Bool;
      "1号梯下行指示" : Bool;
      上行接触器 : Bool;
      下行接触器 : Bool;
      "1层上行呼梯按钮指示灯" : Bool;
      "2层上行呼梯按钮指示灯" : Bool;
      "3层上行呼梯按钮指示灯" : Bool;
      "4层上行呼梯按钮指示灯" : Bool;
      "5层上行呼梯按钮指示灯" : Bool;
      "6层上行呼梯按钮指示灯" : Bool;
      "7层上行呼梯按钮指示灯" : Bool;
      "8层上行呼梯按钮指示灯" : Bool;
      "9层上行呼梯按钮指示灯" : Bool;
      "2层下行呼梯按钮指示灯" : Bool;
      "3层下行呼梯按钮指示灯" : Bool;
      "4层下行呼梯按钮指示灯" : Bool;
      "5层下行呼梯按钮指示灯" : Bool;
      "6层下行呼梯按钮指示灯" : Bool;
      "7层下行呼梯按钮指示灯" : Bool;
      "8层下行呼梯按钮指示灯" : Bool;
      "9层下行呼梯按钮指示灯" : Bool;
      "10层下行呼梯按钮指示灯" : Bool;
      "1号梯1层按钮指示灯" : Bool;
      "1号梯2层按钮指示灯" : Bool;
      "1号梯3层按钮指示灯" : Bool;
      "1号梯4层按钮指示灯" : Bool;
      "1号梯5层按钮指示灯" : Bool;
      "1号梯6层按钮指示灯" : Bool;
      "1号梯7层按钮指示灯" : Bool;
      "1号梯8层按钮指示灯" : Bool;
      "1号梯9层按钮指示灯" : Bool;
      "1号梯10层按钮指示灯" : Bool;
      "1号梯上平层信号" : Bool;
      "1号梯下平层信号" : Bool;
      "1号梯开门到位" : Bool;
      "1号梯关门到位" : Bool;
      正处于故障中 : Bool;
      "存在安全隐患（光幕）" : Bool;
      当前楼层数 : Int;
      "1号梯检修信号" : Bool;
      外呼上面无目标2 : Bool;
      外呼上面无目标3 : Bool;
      外呼上面无目标4 : Bool;
      外呼上面无目标5 : Bool;
      外呼上面无目标6 : Bool;
      外呼上面无目标7 : Bool;
      外呼上面无目标8 : Bool;
      外呼上面无目标9 : Bool;
      外呼下面无目标2 : Bool;
      外呼下面无目标3 : Bool;
      外呼下面无目标4 : Bool;
      外呼下面无目标5 : Bool;
      外呼下面无目标6 : Bool;
      外呼下面无目标7 : Bool;
      外呼下面无目标8 : Bool;
      外呼下面无目标9 : Bool;
      "1号梯轿内开门按钮" : Bool;
      "1号梯轿内关门按钮" : Bool;
      上端站1限位 : Bool;
      下端站1限位 : Bool;
   END_VAR
   VAR_OUTPUT
      "1号梯关门继电器" : Bool;
      "1号梯开门继电器" : Bool;
      "停梯截断(完成关门）" : Bool;
      "停梯截断(完成开门）" : Bool;
      死机 : Bool;
   END_VAR
   VAR
      开门到位次数 : Int;
      开门次数达到上限 : Bool;
      连接46 : Bool;
      连接47 : Bool;
      连接48 : Bool;
      连接49 : Bool;
      连接50 : Bool;
      连接51 : Bool;
      连接52 : Bool;
      连接53 : Bool;
      连接54 : Bool;
      连接55 : Bool;
      连接56 : Bool;
      连接57 : Bool;
      连接58 : Bool;
      连接59 : Bool;
      连接67 : Bool;
      连接68 : Bool;
      连接69 : Bool;
      连接70 : Bool;
      连接71 : Bool;
      连接72 : Bool;
      连接73 : Bool;
      连接74 : Bool;
      连接75 : Bool;
      连接76 : Bool;
      连接77 : Bool;
      连接78 : Bool;
      连接79 : Bool;
      连接80 : Bool;
      连接107 : Bool;
      连接108 : Bool;
      连接109 : Bool;
      连接110 : Bool;
      连接111 : Bool;
      连接112 : Bool;
      连接113 : Bool;
      连接114 : Bool;
      连接115 : Bool;
      连接116 : Bool;
      连接117 : Bool;
      连接118 : Bool;
      连接119 : Bool;
      连接120 : Bool;
      连接121 : Bool;
      连接122 : Bool;
      连接123 : Bool;
      连接124 : Bool;
      连接125 : Bool;
      电梯动过 : Bool;
      分类上行特殊 : Bool;
      分类下行特殊 : Bool;
      完成开门截断 : Bool;
      "0为正常流程，1为非正常" : Bool;
      稍后置零停梯截断完成关门 : TON_TIME;
      保证停梯 : TOF_TIME;
      保证停梯上 : TOF_TIME;
      "稍后置1停梯截断完成关 门" : TON_TIME;
      "保证后面变 量有效置" : TON_TIME;
      "判断 死机" : TON_TIME;
   END_VAR
   VAR RETAIN
      停梯截断开门次数 : CTU_INT;
      判断电梯运动 : CTU_INT;
      计算开门次数 : CTU_INT;
   END_VAR
   VAR
      IEC_Timer_0_Instanc_ : TP_TIME;
      IEC_Timr_0_Instance : TON_TIME;
      IEC_Tim_0_Instance : TON_TIME;
      IEC_Timer_0_Instance : TOF_TIME;
      IEC_Timer_0_Instance_1 : TON_TIME;
   END_VAR
   VAR RETAIN
      计算开门到位次数 : CTU_INT;
   END_VAR
   VAR_TEMP   // added for the SCL form of the ladder/FBD networks
      _w1 : Bool;
      _w2 : Bool;
      _w3 : Bool;
      _w4 : Bool;
      _w5 : Bool;
      _w6 : Bool;
      _w7 : Bool;
      _w8 : Bool;
      _w9 : Bool;
      _w10 : Bool;
      _w11 : Bool;
      _w12 : Bool;
      _w13 : Bool;
      _w14 : Bool;
      _w15 : Bool;
      _w16 : Bool;
      _w17 : Bool;
      _w18 : Bool;
      _w19 : Bool;
      _w20 : Bool;
      _w21 : Bool;
      _w22 : Bool;
   END_VAR
BEGIN

REGION Network 1: 停梯
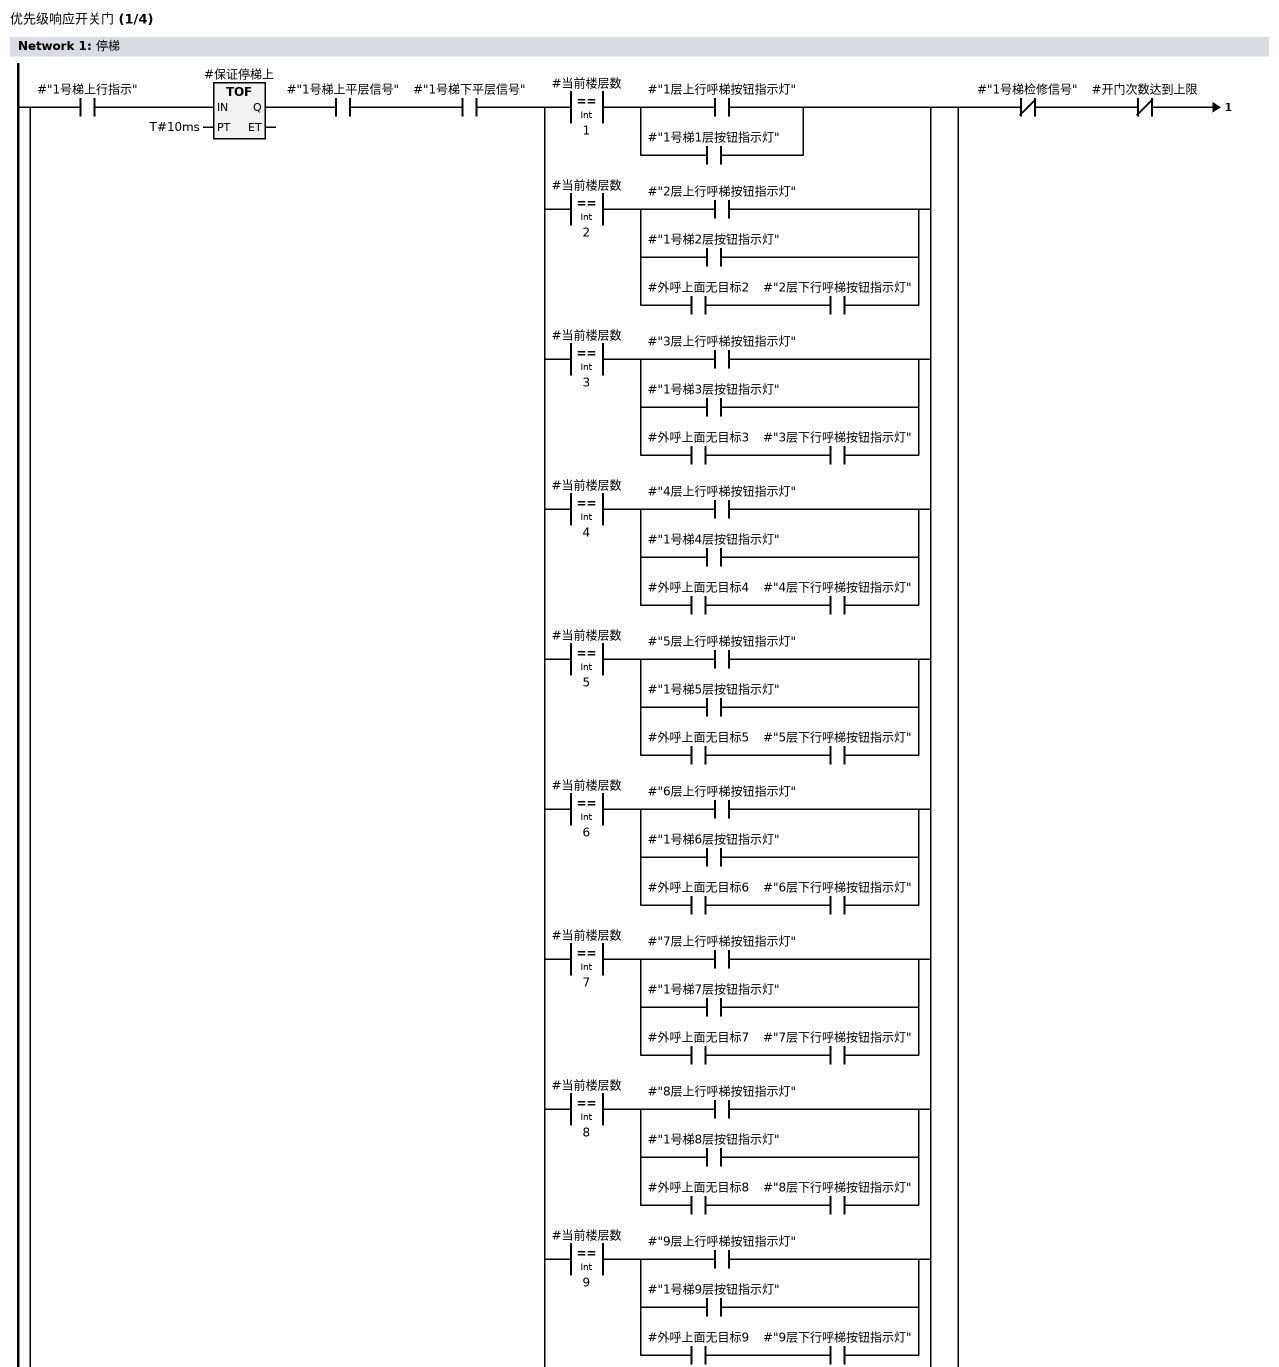
